// I/O API/IN/STRUCTURE/bds_inPha_measmt_ts
///Data structure for one current measurement value of the API function |bds_inPha_get.|.
{attribute 'external_name' := 'cmp_rts_bds_inPha_measmt_ts'}
TYPE bds_inPha_measmt_ts :
STRUCT
	///Measured current in micro Ampere
	phaShift_dDeg_s32 : DINT;
	///Shunt state of the input current measurement signal
	tiPhaDif_ns_u32: UDINT;
	///Measured current in micro Ampere
	tiPerdPrimSig_ns_u32 : UDINT;
	///Shunt state of the input current measurement signal
	tiPerdSecSig_ns_u32: UDINT;
	///Measured current in micro Ampere
	cntPlsPrimSig_u32 : UDINT;
	///Shunt state of the input current measurement signal
	cntPlsSecSig_u32: UDINT;
	///Shunt state of the input current measurement signal
	statusDiag_b: bds_inPha_statusDiag_tb;
	///Status of the measurement
	status_e: bds_inCmn_status_te;
END_STRUCT
END_TYPE

// I/O API/IN/STRUCTURE/bds_inPha_statusDiag_tb
{attribute 'external_name' := 'cmp_rts_bds_inPha_statusDiag_tb'}
{attribute 'size' := '32'}
TYPE bds_inPha_statusDiag_tb :
STRUCT
	stErrPrimSigMaxPerdOvf_b1: BIT; // Fault error status for maximum period overflow on primary signal;
	stErrSecSigMaxPerdOvf_b1: BIT; // Fault error status for maximum period overflow on secondary signal;
	stErrSigFrqMismatch_b1: BIT; // Fault error status for frequency mismatch of primary and secondary signal.
	resd1_b : ARRAY[0..2] OF BYTE;      (* Reserved *)
END_STRUCT
END_TYPE

// I/O API/IN/STRUCTURE/bds_inPha_tiBufdMeasmt_ts
///Data structure for twenty pwm measurement values of the API function |bds_inPwm_getTiBufd|, used to get the buffered values.
{attribute 'external_name' := 'cmp_rts_bds_inPha_tiBufdMeasmt_ts'}
TYPE bds_inPha_tiBufdMeasmt_ts :
STRUCT
	///Up to 20 samples of PWM period in ns, 0th index is latest
	tiPhaDif_ns_au32: ARRAY[0..19] OF UDINT;
	///Up to 20 samples of ON pulse width in ns
	tiPerdPrimSig_ns_au32: ARRAY[0..19] OF UDINT;
	///Up to 20 samples of ON pulse width in ns
	tiPerdSecSig_ns_au32: ARRAY[0..19] OF UDINT;
	///Number of new samples (pulses) received since the last call of API. It is limited to 20 samples.
	cntPlsPrimSig_u32: UDINT;
	///Number of new samples (pulses) received since the last call of API. It is limited to 20 samples.
	cntPlsSecSig_u32: UDINT;
	///Number of new samples (pulses) received since the last call of API. It is limited to 20 samples.
	cntNewSample_u32: UDINT;
	///Number of new samples (pulses) received since the last call of API. It is limited to 20 samples.
	statusDiag_b: bds_inPha_statusDiag_tb;
END_STRUCT
END_TYPE

// I/O API/IN/STRUCTURE/bds_inPha_tiBufd_ts
///Data structure for pwm measurement value of the API function |bds_inPha_tiBufd_ts|.
{attribute 'external_name' := 'cmp_rts_bds_inPha_tiBufd_ts'}
TYPE bds_inPha_tiBufd_ts :
STRUCT
	///Status of the measurement
	status_e: bds_inCmn_status_te;
END_STRUCT
END_TYPE

// System API/DSM/DSM Refactored( 3-byte DTC)/STRUCTURE/bds_dsmCmn_stWord_tb
///Structure for the Bit field for the 16-bit status word of DFC.
{attribute 'external_name' := 'cmp_rts_bds_dsmCmn_stWord_tb'}
TYPE bds_dsmCmn_stWord_tb :
STRUCT
	///Fault level (0x0 - OK level, 0xF - Defect)
	stFltLvl_b4: BIT;
	///Status of Last Debounced Fault (LDF)
	stLDF_b1: BIT;
	///Tested Since Clear Status (1 - Yes, 0 - No)
	stTSC_b1: BIT;
	///Memory Status (DFC is saved in fault memory or not)
	stMS_b1: BIT;
	///Debounce Active Status (1 - Yes, 0 - No)
	stDA_b1: BIT;
	///Debounced Fault Level (With five levels 0x0, 0x4, 0x8, 0xC and 0xF (e.g., 0xC = 75% debounced)
	stDebdFltLvl_b4: BIT;
	///Fault Since Clear Status (1=Yes, 0=No)
	stFSC_b1: BIT;
	///Test Status
	stTestSt_b1: BIT;
	///Not used
	stUnused_b1: BIT;
	///Test finalized
	stNotFinalized_b1: BIT;
END_STRUCT
END_TYPE

// System API/DSM/DSM Refactored( 3-byte DTC)/STRUCTURE/bds_dsmDTC_deleteErr_ts
///Return structure for bds_dsmDTC_deleteErr POU.
{attribute 'external_name' := 'cmp_rts_bds_dsmDTC_deleteErr_ts'}
TYPE bds_dsmDTC_deleteErr_ts :
STRUCT
	///Status or result of POU operation 
	apiSt_e: bds_dsmCmn_st_te;
END_STRUCT
END_TYPE

// System API/DSM/DSM Refactored( 3-byte DTC)/STRUCTURE/bds_dsmDTC_getDFES_ts
///Return structure for bds_dsmDTC_getDFES POU.
{attribute 'external_name' := 'cmp_rts_bds_dsmDTC_getDFES_ts'}
TYPE bds_dsmDTC_getDFES_ts :
STRUCT
	///Number of errors returned
	nrErr_u8: USINT;
	///DTCs as in DFES array
	dtcListDFES_au32: ARRAY[1..32] OF UDINT;
	///Status or result of POU operation (Valid POU call / Invalid parameter (invalid mask)/ out of Range (DTC value out of range)) 
	apiSt_e: bds_dsmCmn_st_te;
END_STRUCT
END_TYPE

// System API/DSM/DSM Refactored( 3-byte DTC)/STRUCTURE/bds_dsmDTC_getDTCVal_ts
///Return structure for bds_dsmDTC_getDTCVal POU.
{attribute 'external_name' := 'cmp_rts_bds_dsmDTC_getDTCVal_ts'}
TYPE bds_dsmDTC_getDTCVal_ts :
STRUCT
	///DTC value
	dtc_u32: UDINT;
	///Status or result of API operation (API call successful / invalid config (wrong DFC passed) 
	apiSt_e: bds_dsmCmn_st_te;
END_STRUCT
END_TYPE

// System API/DSM/DSM Refactored( 3-byte DTC)/STRUCTURE/bds_dsmDTC_getErrList_ts
///Return structure for bds_dsmDTC_getErrList POU.
{attribute 'external_name' := 'cmp_rts_bds_dsmDTC_getErrList_ts'}
TYPE bds_dsmDTC_getErrList_ts :
STRUCT
	///Number of errors returned
	nrErr_u8: USINT;
	///DTC list containing 32 entries
	dtcList_au32: ARRAY[1..32] OF UDINT;
	///Status or result of POU operation (Valid POU call / Invalid parameter (invalid mask) 
	apiSt_e: bds_dsmCmn_st_te;
END_STRUCT
END_TYPE

// System API/DSM/DSM Refactored( 3-byte DTC)/STRUCTURE/bds_dsmDTC_getStatus_ts
///Return structure for bds_dsmDTC_getStatus POU.
{attribute 'external_name' := 'cmp_rts_bds_dsmDTC_getStatus_ts'}
TYPE bds_dsmDTC_getStatus_ts :
STRUCT
	///Error State (Active / Previously Active / Deactive)
	errState_e: UDINT;
	///DTC Detailed Status Parameters as 16 bit Status Word in DFC
	stWordDTC_b: bds_dsmCmn_stWord_tb;
	///Status or result of POU operation 
	apiSt_e: bds_dsmCmn_st_te;
END_STRUCT
END_TYPE

// System API/DSM/DSM Refactored( 3-byte DTC)/STRUCTURE/bds_dsmDTC_updateErr_ts
///Return structure for bds_dsmDTC_updateErr POU.
{attribute 'external_name' := 'cmp_rts_bds_dsmDTC_updateErr_ts'}
TYPE bds_dsmDTC_updateErr_ts :
STRUCT
	///Status or result of POU operation
	apiSt_e: bds_dsmCmn_st_te;
END_STRUCT
END_TYPE

// Communication API/ISOBUS/J1939-76/STRUCTURE/bds_isobus_cnsrDataboxInfo_ts
///Structure of the consumer data box information
{attribute 'external_name' := 'cmp_rts_bds_isobus_cnsrDataboxInfo_ts'}
TYPE bds_isobus_cnsrDataboxInfo_ts :
STRUCT
	///pointer to the consumer SDG databox buffer
	mem_pas: POINTER TO bds_isobus_cnsrSdgMsg_ts;
	///number of SDG messages to be received
	numOfMsg_u16: UINT;
END_STRUCT
END_TYPE

// Communication API/ISOBUS/J1939-76/STRUCTURE/bds_isobus_cnsrSdgMsg_ts
///Structure for handling Consumer databox
{attribute 'external_name' := 'cmp_rts_bds_isobus_cnsrSdgMsg_ts'}
TYPE bds_isobus_cnsrSdgMsg_ts :
STRUCT
	///pointer to data array with length=lenMax_u8
	data_pau8: POINTER TO USINT;
	///function is called if SDG is received and processed
	func_pf: POINTER TO UINT;
	///CAN Id of the SDM to be received
	canID_u: bds_isobus_sfty_canID_tu;
	///length of received SDM message
	lenAct_u8: USINT;
	///max length of the SDG receive buffer defined
	lenMax_u8: USINT;
	///expected maximum time between consecutive SDMs received
	sct_u32: UDINT;
	///expected maximum time between SHM and SDM of an SDG received
	srvt_u32: UDINT;
	///expected Source address of the sender (i.e., Producer)
	srcAddr_u8: USINT;
	///status of consumer SDG databox
	status_u16: UINT;
	///flag to identify first message received after start-up
	firstSdg_l: BOOL;
	///SCT timer
	sctTmr_s: bds_isobus_sftyTmr_ts;
	///SRVT timer
	srvtTmr_s: bds_isobus_sftyTmr_ts;
	///SDM CRC
	sdmCrc_u: bds_isobus_sdmCrcVal_tu;
	///sequence number handling structure
	seqNum_s: bds_isobus_cnsrSdgSeqNum_ts;
	///SDG state handling enumeration
	sdgState_e: bds_isobus_sdgState_te;
	///Status of Consumer to be updated to ASW
	cnsrStatus_e: bds_isobus_sdgCnsrStatus_te;
END_STRUCT
END_TYPE

// Communication API/ISOBUS/J1939-76/STRUCTURE/bds_isobus_cnsrSdgSeqNum_ts
///Structure type definition for handling CRC32 value of SDM
{attribute 'external_name' := 'cmp_rts_bds_isobus_cnsrSdgSeqNum_ts'}
TYPE bds_isobus_cnsrSdgSeqNum_ts :
STRUCT
	///Sequence number of currently received SDG
	curSdgSeqNum_u8: UINT;
	///Sequence number of previously received SDG, initialize with 0xFF to monitor 0th sequence after start-up
	prevSdgSeqNum_u8: UINT;
END_STRUCT
END_TYPE

// Communication API/ISOBUS/J1939-76/STRUCTURE/bds_isobus_prodDataboxInfo_ts
///Structure of the producer data box information
{attribute 'external_name' := 'cmp_rts_bds_isobus_prodDataboxInfo_ts'}
TYPE bds_isobus_prodDataboxInfo_ts :
STRUCT
	///pointer to the consumer SDG databox buffer
	mem_pas: POINTER TO bds_isobus_prodSdgMsg_ts;
	///number of SDG messages to be transmitted
	numOfMsg_u16: UINT;
END_STRUCT
END_TYPE

// Communication API/ISOBUS/J1939-76/STRUCTURE/bds_isobus_prodSdgMsg_ts
///Structure for handling Producer databox
{attribute 'external_name' := 'cmp_rts_bds_isobus_prodSdgMsg_ts'}
TYPE bds_isobus_prodSdgMsg_ts :
STRUCT
	///pointer to data array updated in Producer callback with length=lenMax_u8
	data_pau8: POINTER TO USINT;
	///function is called before SDG is to be sent (Producer Callback)
	func_pf: POINTER TO UINT;
	///CAN Id of the SDM to be sent
	canID_u: bds_isobus_sfty_canID_tu;
	///max length (buffer size) of SDM to be sent
	lenMax_u8: USINT;
	///actual length of SDM message to be sent
	lenAct_u8: USINT;
	///cycle time for fixed transmission of the SDG
	cycle_u16: UINT;
	///counter for monitoring cyclic transmission of SDG
	counter_u16: UINT;
	///expected Source address of the sender (i.e., Producer)
	srcAddr_u8: USINT;
	///status of Producer SDG databox
	status_u16: UINT;
	///Databox number of the SDG being handled
	SdgDataboxNum_u16: UINT;
	///SDM CRC
	sdmCrc_u: bds_isobus_sdmCrcVal_tu;
	///Sequence number of the SDG being handled
	seqNum_u8: USINT;
	///Timer value of previously transmitted SDG //ToDo: for variable transmission
	prevSdgTmrVal_u32: UDINT;
	///Structure instance containing SHM related data
	shmMsg_s: bds_isobus_shmMsg_ts;
END_STRUCT
END_TYPE

// Communication API/ISOBUS/J1939-76/UNION/bds_isobus_sdmCrcVal_tu
///Union type definition for handling CRC32 value of SDM
{attribute 'external_name' := 'cmp_rts_bds_isobus_sdmCrcVal_tu'}
TYPE bds_isobus_sdmCrcVal_tu :

UNION
	///array containing CRC32 data bytes
	sdmCrcVal_au8: ARRAY[1..4] OF USINT;
	///CRC32 value
	sdmCrcVal_u32: UDINT;
END_UNION

END_TYPE

// Communication API/ISOBUS/J1939-76/STRUCTURE/bds_isobus_sftyTmr_ts
///Structure type definition for Timer handling
{attribute 'external_name' := 'cmp_rts_bds_isobus_sftyTmr_ts_ts'}
TYPE bds_isobus_sftyTmr_ts :
STRUCT
	///timer value for monitoring
	tmrStrd_u32: UDINT;
END_STRUCT
END_TYPE

// Communication API/ISOBUS/J1939-76/STRUCTURE/bds_isobus_sfty_canID_ts
///Structure for handling CAN Id of SHM and SDM.
{attribute 'external_name' := 'cmp_rts_bds_isobus_sfty_canID_ts'}
TYPE bds_isobus_sfty_canID_ts :
STRUCT
	/// node id of the transmitter 
	SourceAddr_b8: BYTE;
	/// if PF<240, this value is destination address else Group extension
	PDUSpecific_b8: BYTE;
	/// this byte determines whether the message can be transmitted with a destination address or as a broadcast
	PDUFormat_b8: BYTE;
	/// these bits identify the data pages of the parameter group
	DataPage_b2: BIT;
	/// these 3 bits define the priority of the following message
	Priority_b3: BIT;
	/// these 3 bits are overhead for the 29 bit CAN Id 
	unusedBits_b3: BIT;
END_STRUCT
END_TYPE

// Communication API/ISOBUS/J1939-76/UNION/bds_isobus_sfty_canID_tu
///Union type definition for handling CAN Id of SHM and SDM
{attribute 'external_name' := 'cmp_rts_bds_isobus_sfty_canID_tu'}
TYPE bds_isobus_sfty_canID_tu :

UNION
	///CAN Id structure of type bds_isobus_sfty_canID_ts
	canID_s: bds_isobus_sfty_canID_ts;
	///CAN Id value
	canID_u32: UDINT;
END_UNION

END_TYPE

// Communication API/ISOBUS/J1939-76/STRUCTURE/bds_isobus_shmMsg_ts
///Structure containing SHM parameters of the bds_isobus_prodSdgMsg_t SDG databox being handled
{attribute 'external_name' := 'cmp_rts_bds_isobus_shmMsg_ts'}
TYPE bds_isobus_shmMsg_ts :
STRUCT
	///array containing CRC32 data bytes
	data_au8: ARRAY[1..8] OF USINT;
	///CAN Id of the SDM to be received
	canID_u: bds_isobus_sfty_canID_tu;
END_STRUCT
END_TYPE

// System API/DSM/DSM Refactored( 3-byte DTC)/ENUM/bds_dsmCmn_st_te
(* common status enumeration return types*)
{attribute 'external_name' := 'cmp_rts_bds_dsmCmn_st_te'}
TYPE bds_dsmCmn_st_te :
(
	(*POU call successful*)
	bds_dsmCmn_ok_E := 0,
	(*Parameter out of Range (e.g., invalid DTC value, which is not within the configured Range)*)
	bds_dsmCmn_outOfRng_E,
	(*not available (e.g. busy, called to early in init, System in a mode it cannot measure etc.)*)
    bds_dsmCmn_notAvl_E,
	(*POU call invalid, e.g., calling a not configured DFC, etc.*)
    bds_dsmCmn_invldCfg_E,
	(*POU call invalid because of invalid Parameter*)
    bds_dsmCmn_invldPrm_E,
	(*POU call invalid because of invalid pointer*)
    bds_dsmCmn_invldPtr_E,
	(*Not available due to an internal error*)
    bds_dsmCmn_errInt_E
	
)USINT;
END_TYPE

// System API/DSM/DSM Refactored( 3-byte DTC)/ENUM/bds_dsmCmn_errState_te
(*Enumeration containing the error state of DFC (Active / Previously Active / Deactive).*)
{attribute 'external_name' := 'cmp_rts_bds_dsmCmn_errState_te'}
TYPE bds_dsmCmn_errState_te :
(
	(*Error is Active*)
	bds_dsmCmn_stErrActv_e := 1,
	(*Error is Previously Active*)
	bds_dsmCmn_stErrPrevActv_e,
	(*Error is in Deactive State*)
	bds_dsmCmn_stErrDeactv_e
	
)USINT;
END_TYPE

// System API/DSM/DSM Refactored( 3-byte DTC)/ENUM/bds_dsmCmn_fltLvl_te
(*Enumeration for fault level of a DFC, as a result of check.*)
{attribute 'external_name' := 'cmp_rts_bds_dsmCmn_fltLvl_te'}
TYPE bds_dsmCmn_fltLvl_te :
(
	(*Fault percent 0%*)
	bds_dsmCmn_fltLvl_0_Perc_e := 0,
	(*Fault percent 100%*)
	bds_dsmCmn_fltLvl_100_Perc_e
	
)USINT;
END_TYPE

// System API/DSM/DSM Refactored( 3-byte DTC)/STRUCTURE/bds_dsmJ1939_LampSt_tb
(*Bit field for Lamp States.*)
{attribute 'external_name' := 'cmp_rts_bds_dsmJ1939_LampSt_tb'}
TYPE bds_dsmJ1939_LampSt_tb :
STRUCT
	(*Lamp/Flash State of Malfunction Indicator Lamp (MIL)*)
	milSt_b2: BIT;
	(*Lamp/Flash State of Red Stop Lamp (RSL)*)
	rslSt_b2: BIT;
	(*Lamp/Flash State of Amber Warning Lamp (AWL)*)
	awlSt_b2: BIT;
	(*Lamp/Flash State of Protected Lamp (PRL)*)
	prlSt_b2: BIT;
END_STRUCT
END_TYPE

// System API/DSM/DSM Refactored( 3-byte DTC)/STRUCTURE/bds_dsmJ1939_getJ1939DTC_ts
(*Return structure for the bds_dsmJ1939_getJ1939DTC POU.*)
{attribute 'external_name' := 'cmp_rts_bds_dsmJ1939_getJ1939DTC_ts'}
TYPE bds_dsmJ1939_getJ1939DTC_ts :
STRUCT
	(*SPN value*)
	spn_u32 : UDINT;
	(*FMI value*)
	fmi_u8 : USINT;
	(*Bitfield containing Lamp States (MIL, RSL, AWL, Protected Lamp)*)
	lampSt_b : bds_dsmJ1939_LampSt_tb;
	(*Occurrence Counter*)
	occCntr_u8 : USINT;
	(* Status or result of POU operation (Valid POU call / DTC passed is out of range)*)
	apiSt_e : bds_dsmCmn_st_te;
END_STRUCT
END_TYPE

// Communication API/CAN/CAN-FD legacy/ENUM/bds_can_fd_St_te
{attribute 'external_name' := 'cmp_rts_bds_can_fd_St_te'}
TYPE bds_can_fd_St_te :
(
	//API call successful
    bds_can_fd_ok_E := 0,
	//Databox not empty
    bds_can_fd_txDataboxNotEmpty_E := 1,
	//Invalid Access to FFI variant API call.
    bds_can_fd_errFfi_E := 5,
	//Invalid CAN-FD databox number
    bds_can_fd_invldDataBoxNbr_E := 9,
	//Invalid CAN-FD channel
    bds_can_fd_invldChnl_E := 14,
	//Invalid CAN-FD identifier
    bds_can_fd_invldId_E := 15,
	//Invalid CAN-FD message format
    bds_can_fd_invldFormat_E := 16,
	//Invalid number of bytes
    bds_can_fd_invldNumBytes_E := 17,
	//Number of messages registered in buffer = 0
    bds_can_fd_numMsgZero_E := 18,
	//CAN-FD transmit buffer overflow
    bds_can_fd_txBufOvfl_E := 20,
	//CAN-FD receive buffer overflow
    bds_can_fd_rxBufOvfl_E := 30,
	//CAN-FD receive buffer is empty
    bds_can_fd_rxBufEmpty_E := 31,
	//CAN-FD receive buffer length is zero
    bds_can_fd_rxBufLenZero_E := 32,
	//Buffer address overlap
    bds_can_fd_ovlpAddr_E := 55,
	//Invalid address
    bds_can_fd_invldAddr_E := 60,
	//Invalid address (parameter buf_pas). Buffer length is zero
    bds_can_fd_rxDataboxBufLenZero_E := 61,
	//Databox not initialized
    bds_can_fd_dataBoxNoInit_E := 62,
	//Databox with this identifier is initialized already, new initialization is not accepted
    bds_can_fd_errDataboxIdExist_E := 63,
	//Number of databoxes registered is greater than previously registered number of databoxes
    bds_can_fd_prevRegdDataboxMoreThanCurrent_E := 64,
	//Invalid number of databoxes
    bds_can_fd_invldCfgDatabox_E := 65,
	//CAN hardware not supported in RC.
    //e.g., 3 CAN channel RC5-6/40 ECU.
    bds_can_fd_hwNotSupported_E := 66,
	//Configuration not allowed
    bds_can_fd_cfgNotAllowed_E := 99,
	//CAN-FD not supported in CAN_3
    bds_can_fd_paramChnl3Err_E := 100
)USINT;
END_TYPE

// Communication API/CAN/CAN-FD legacy/STRUCTURE/bds_can_fd_Message_ts
{attribute 'external_name' := 'cmp_rts_bds_can_fd_Message_ts'}
TYPE bds_can_fd_Message_ts :
STRUCT
	//Identifier of the message.
	//Value range:
	// 16#000 .. 0x7FF (11-bit standard format)
	// 16#00000000 .. 0x1FFFFFFF (29-bit extented format)
	id_u32 : UDINT;
	//Format of the CAN-FD message.Value range:
    //BDS_CAN_STD_DU8 (11-bit standard format)
	//BDS_CAN_EXD_DU8 (29-bit extented format)
	format_u8 : USINT;
	//Number of data bytes which will be transmitted or which type received.
	numBytes_u8 : USINT;
	//Data which will be transmitted or which were received.Size of the define, bds_can_fd_maxDataBytes_DU8 is equal to 64.
	data_au8 : ARRAY[0..63] OF USINT;
END_STRUCT
END_TYPE

// Communication API/ISOBUS/J1939-76/ENUM/bds_isobus_sdgCnsrStatus_te
(*Enumeration for Consumer SDG reception status.*)
{attribute 'external_name' := 'cmp_rts_bds_isobus_sdgCnsrStatus_te'} 
TYPE  bds_isobus_sdgCnsrStatus_te :
(  
	(*valid SDG received*)
	bds_isobus_sdgCnsrOk_E := 0,
	(*SRVT timeout*)
	bds_isobus_sdgCnsrSrvtTmngErr_E,
	(*SCT timeout*)
	bds_isobus_sdgCnsrSctTmngErr_E,
	(*SDG received with invalid CRC*)
    bds_isobus_sdgCnsrCrcError_E,
	(*SDG received with invalid sequence number*)
    bds_isobus_sdgCnsrSeqError_E,
	(*SDG received with invalid data length*)
    bds_isobus_sdgCnsrLenError_E
)USINT;
END_TYPE

// Communication API/ISOBUS/J1939-76/ENUM/bds_isobus_sdgState_te
(*Enumeration for Consumer SDG reception status.*)
{attribute 'external_name' := 'cmp_rts_bds_isobus_sdgState_te'} 
TYPE bds_isobus_sdgState_te :
(
	(*SDG initialized*)
	bds_isobus_sfty_sdgIniDone_E := 0,
	(*SHM received and processed*)
	bds_isobus_sfty_shmProcessed_E,
	(*both SHM and SDM received and processed*)
	bds_isobus_sfty_sdgProcessed_E,
	(*SRVT timeout*)
	bds_isobus_sfty_srvtExpired_E,
	(*SCT timeout*)
	bds_isobus_sfty_sctExpired_E,
	(*SDG successfully validated*)
	bds_isobus_sfty_sdgValidated_E,
	(*Consumer SDG callback triggered*)
	bds_isobus_sfty_cnsrSdgCbkTriggered_E
)USINT;
END_TYPE

// Communication API/ISOBUS/J1939-76/ENUM/bds_isobus_sfty_apiRetVal_te
(*Enumeration for J1939-76 API return values.*)
{attribute 'external_name' := 'cmp_rts_bds_isobus_sfty_apiRetVal_te'}
TYPE bds_isobus_sfty_apiRetVal_te :
(
	(*No API execution error*)
	 bds_isobus_sfty_noErr_E := 0,
	(*invalid address*)
	 bds_isobus_sfty_invldAdr_E,
	(*address overlaps with other buffers*)
 	 bds_isobus_sfty_ovlAdr_E,
	(*invalid CA instance number*)
	 bds_isobus_sfty_invldInstNum_E,
	(*message box is not yet initialized*)
	 bds_isobus_sfty_boxStNoIni_E,
	(*configuration is not allowed*)
	 bds_isobus_sfty_boxStIni_E,
	(*invalid databox number*)
	 bds_isobus_sfty_cfgNotAllwd_E,
	(*invalid PGN value*)
	 bds_isobus_sfty_invldDataboxNum_E,
	(* invalid priority of SDG*) 
	 bds_isobus_sfty_invldPgn_E,
	(*invalid cycle time for SDG*)
	 bds_isobus_sfty_invldPrio_E,
	(*invalid offset time for SDG*)
	 bds_isobus_sfty_invldCyc_E,
	(*invalid data length of SDM*)
	 bds_isobus_sfty_invldOffs_E,
	(*invalid data address*)
	 bds_isobus_sfty_invldDataLen_E,
	(*Another data box with this id was initialized already*) 
	 bds_isobus_sfty_invldDataPtr_E,
	(*sdg databox initialized*) 
	 bds_isobus_sfty_pgnPrioExists_E,
	(*invalid source address*)
	 bds_isobus_sfty_invldSrcAdr_E,
	(*invalid SCT*)
	 bds_isobus_sfty_invldSct_E,
	(*invalid SRVT*) 
	 bds_isobus_sfty_invldSrvt_E,
	(*Internal PGN used*) 
	 bds_isobus_sfty_intPgnUsed_E,
	(*API used without enabling J1939-76 feature in eC*)
	 bds_isobus_sfty_featNotEnad_E,
	(*Invalid pointer*)
	 bds_isobus_sfty_invldCbkAdr_E
)USINT;
END_TYPE

// Diagnostics API/UDS/ENUM/bds_udsCmn_statusApi_te
{attribute 'external_name' := 'cmp_rts_bds_udsCmn_statusApi_te'}
TYPE bds_udsCmn_statusApi_te :
(
	(*Success: API executed without error*)
	bds_udsCmn_ok_E := 0,
	(*Invalid: calling an unconfigured signal/DID *)
	bds_udsCmn_invldCfg_E,
	(*Invalid: invalid parameter*)
	bds_udsCmn_invldPrm_E,
	(*Out of range: the array size should be less than or equal to 17 bytes*)
	bds_udsCmn_outOfRng_E,
	(*not available: (e.g. busy, called to early in init, system is in a mode that it cannot measure etc)*)
	bds_udsCmn_notAvl_E
)USINT;
END_TYPE

// Communication API/CAN/CAN-FD legacy/STRUCTURE/bds_can_fd_RxDatabox_ts
///Structure of a CAN-FD receive (Rx) databox.
{attribute 'external_name' := 'cmp_rts_bds_can_fd_RxDatabox_ts'}
TYPE bds_can_fd_RxDatabox_ts :
STRUCT
	//CAN ID
    //Value range:
    //16#000 .. 0x7FF (11-bit standard format)
    // 16#00000000 .. 16#1FFFFFFF (29-bit extented format)
	id_u32 : UDINT;
	//CAN ID format
    //Value range:
    //BDS_CAN_STD_DU8 (11-bit standard format)
    //BDS_CAN_EXD_DU8 (29-bit extented format)
	format_u8 : USINT;
	//Number of data bytes which will be received.
    numBytes_u8 : USINT;
	//Pointer to callback function for CAN-FD Receive Databox
    callback_pf : UINT;
	//Structure instance to CAN-FD databox buffer information
    Buf_s : bds_can_fd_DataboxBufInfo_ts;
END_STRUCT
END_TYPE

// Communication API/CAN/CAN-FD legacy/STRUCTURE/bds_can_fd_DataboxData_ts
///Structure of data of a CAN-FD databox.
{attribute 'external_name' := 'cmp_rts_bds_can_fd_DataboxData_ts'}
TYPE bds_can_fd_DataboxData_ts :
STRUCT
	//Received data.Size of the define, bds_can_fd_maxDataBytes_DU8 is equal to 64.
	data_au8 : ARRAY[0..63] OF USINT;
	//Number of data bytes received
	numBytes_u8 : USINT;
END_STRUCT
END_TYPE

// Communication API/CAN/CAN-FD legacy/STRUCTURE/bds_can_fd_DataboxBufInfo_ts
///Structure for a CAN-FD databox buffer. Only data of the CAN-FD message is buffered.
{attribute 'external_name' := 'cmp_rts_bds_can_fd_DataboxBufInfo_ts'}
TYPE bds_can_fd_DataboxBufInfo_ts :
STRUCT
	//Pointer to structure for CAN-FD Databox Data structure.
	start_pas : POINTER TO bds_can_fd_DataboxData_ts;
	//CAN-FD Databox Buffer Management Structure 
	Manage_s : bds_can_fd_BufManage_ts;
END_STRUCT
END_TYPE

// Communication API/CAN/CAN-FD legacy/STRUCTURE/bds_can_fd_BufManage_ts
///Structure for a CAN-FD Message Buffer Management.
{attribute 'external_name' := 'cmp_rts_bds_can_fd_BufManage_ts'}
TYPE bds_can_fd_BufManage_ts :
STRUCT
	//Length of the buffer
	length_u16 : UINT;
	//Index for write (CAN-FD send / receive) in the buffer.This is for buffer (FIFO - in sequence value).
	//This is more specific to BSW, has lesser significance to application.
	idx_in_u16 : UINT;
	//Index for read (CAN-FD send / receive) out of the buffer.This is for buffer ((FIFO - out sequence value).
	//This is more specific to BSW, has lesser significance to application.
    idx_out_u16 : UINT;
	//FALSE: Buffer is not empty. If then idx_out - idx_in: buffer is full (no put in).
    //TRUE: Buffer is empty (nothing is to send or nothing was received)
	BufEmpty_l : BOOL;
	//This flag shows if a buffer overflow is occurred.
	//FALSE: No buffer overflow is occurred since last user inquiry of status
    //TRUE: Buffer overflow is occurred.
    BufOvfl_l : BOOL;
END_STRUCT
END_TYPE

// Communication API/CAN/CAN-FD legacy/STRUCTURE/bds_can_fd_TxDatabox_ts
///Structure of a CAN-FD transmit (Tx) databox.
{attribute 'external_name' := 'cmp_rts_bds_can_fd_TxDatabox_ts'}
TYPE bds_can_fd_TxDatabox_ts :
STRUCT
	//CAN ID
    //Value range:
    //16#000 .. 0x7FF (11-bit standard format)
    // 16#00000000 .. 16#1FFFFFFF (29-bit extented format)
	id_u32 : UDINT;
	//CAN ID format
    //Value range:
    //BDS_CAN_STD_DU8 (11-bit standard format)
    //BDS_CAN_EXD_DU8 (29-bit extented format)
	format_u8 : USINT;
	//Number of data bytes which will be received.
    numBytes_u8 : USINT;
	//Data which will be transmitted or which were received.Size of the define, bds_can_fd_maxDataBytes_DU8 is equal to 64.
	data_au8 : ARRAY[0..63] OF USINT;
	//TRUE = databox is empty
    //FALSE = databox contains data which were not sent
    empty_l : BOOL;
	//TRUE = databox is initialized
    //FALSE = databox is not yet initialized
    init_l : BOOL;
END_STRUCT
END_TYPE

// Communication API/ISOBUS/STRUCTURE/bds_isobus_caAddrInfoTbl_ts
///Structure definition of an ISOBUS address info table.
{attribute 'external_name' := 'cmp_rts_bds_isobus_caAddrInfoTbl_ts'}
TYPE bds_isobus_caAddrInfoTbl_ts :
STRUCT
	//ISOBUS CA Name, which is 8 bytes in size according to the ISOBUS/J1939 specification.
	caName_au8 : ARRAY[0..7] OF USINT;
	//ISOBUS CA address which is 1 byte in size.
	caAddr_u8 : USINT;
END_STRUCT
END_TYPE

// Diagnostics API/UDS/STRUCTURE/bds_uds_getActiveService_ts
///Return structure for the API function bds_uds_getActiveService.
{attribute 'external_name' := 'cmp_rts_bds_uds_getActiveService_ts'}
TYPE bds_uds_getActiveService_ts :
STRUCT
	//Status of the UDS API function call.
	stsApi_e : bds_udsCmn_statusApi_te;
	//The value of the UDS service identifier.
    dataSid_u8 : USINT;
END_STRUCT
END_TYPE

// Communication API/ISOBUS/ENUM/bds_isobus_caAddrCbEventType_te
{attribute 'external_name' := 'cmp_rts_bds_isobus_caAddrCbEventType_te'}
TYPE bds_isobus_caAddrCbEventType_te :
(
	//Address claim message received, address table entry is not updated
	bds_isobus_addrClaimMsgRcv_E := 0,
	//Address claim message received and address table entry is updated with new address
    bds_isobus_caTbleAddressUpdate_E,
	//Address claim message received and new entry created in address table
	bds_isobus_caTbleNewEntry_E
)USINT;
END_TYPE

// Communication API/ISOBUS/STRUCTURE/bds_isobus_caAddrInfoTblRef_ts
//Structure type definition to hold reference to Address table info and size of address table info
{attribute 'external_name' := 'cmp_rts_bds_isobus_caAddrInfoTblRef_ts'}
TYPE bds_isobus_caAddrInfoTblRef_ts :
STRUCT
	//pointer to Address Info table
	mem_pas : POINTER TO bds_isobus_caAddrInfoTbl_ts;
	//Total number (Size) of Entries in address info table
	numOfEntry_u8 : USINT;
	//Last valid entry/Number of valid entries in address info table
	lastEntry_u8 : USINT;
END_STRUCT
END_TYPE

// Communication API/Ethernet/STRUCTURE/bds_ethIPv4_getLocalIpAdr_ts
{attribute 'external_name' := 'cmp_rts_bds_ethIPv4_getLocalIpAdr_ts'}
TYPE bds_ethIPv4_getLocalIpAdr_ts :
STRUCT
	//The return structure containing the status information
	statusApi_e : bds_ethIPv4_statusApi_te; 
END_STRUCT
END_TYPE

// Communication API/Ethernet/ENUMS/bds_ethIPv4_statusApi_te
{attribute 'external_name' := 'cmp_rts_bds_ethIPv4_statusApi_te'}
TYPE bds_ethIPv4_statusApi_te :
(
	//API call is successful
	bds_ethIPv4_Adr_Mask_ok_E := 0,
	//API call is invalid because of invalid IPv4 address
    bds_ethIPv4_Adr_Nok_E := 1,
	//API call is invalid because of invalid subnet mask, subnet mask should be 16
    bds_ethIPv4_Mask_Nok_E := 2,
	//Not Available (e.g. busy, called too early in init, not called from OsIniProc etc.)
    bds_ethIPv4_Api_NotAvailable_E := 3, 
	//Invalid parameter passed
    bds_ethIPv4_NullPtr_E := 4, 
    bds_ethIPv4_notAssigned_E :=5 
)USINT;
END_TYPE

// Communication API/Ethernet/STRUCTURE/bds_ethIPv4_setLocalIpAdr_ts
{attribute 'external_name' := 'cmp_rts_bds_ethIPv4_setLocalIpAdr_ts'}
TYPE bds_ethIPv4_setLocalIpAdr_ts :
STRUCT
	//The return structure containing the status information
	statusApi_e : bds_ethIPv4_statusApi_te; 
END_STRUCT
END_TYPE

// Communication API/Ethernet/STRUCTURE/bds_ethIPv4_LocalIpAdr_ts
//Data Structure for IPv4 Address and Subnet Mask for Ethernet functions - bds_ethIPv4_setLocalIpAdr and bds_ethIPv4_getLocalIpAdr
{attribute 'external_name' := 'cmp_rts_bds_ethIPv4_LocalIpAdr_ts'}
TYPE bds_ethIPv4_LocalIpAdr_ts :
STRUCT
	//4 bytes of IPv4 Address
	Ipv4Adr_u32 : UDINT;
	//1 byte of Subnet Mask for IPv4
	Ipv4SubnetMask_u8 : USINT;
END_STRUCT
END_TYPE

// Communication API/Ethernet/ENUMS/bds_ethIPv4_linkState_te
//This enum defines the return values for API bds_ethIPv4_setDoipAdr.
{attribute 'external_name' := 'cmp_rts_bds_ethIPv4_linkState_te'}
TYPE bds_ethIPv4_linkState_te :
(
	bds_ethIPv4_linkDown_E := 0,
	bds_ethIPv4_linkUp_E := 1,
	bds_ethIPv4_linkUndef_E
)USINT;
END_TYPE

// Communication API/Ethernet/ENUMS/bds_ethIPv4_retDoipAdr_te
//This enum defines the return values for API bds_ethIPv4_setDoipAdr.
{attribute 'external_name' := 'cmp_rts_bds_ethIPv4_retDoipAdr_te'}
TYPE bds_ethIPv4_retDoipAdr_te :
(
	//Address set successfully 
	bds_ethIPv4_retAdrOk_E := 0,
	//RC4x Logical Address out of range
	bds_ethIPv4_retLogAdrNok_E :=1,
	//Tester Address out of range
	bds_ethIPv4_retTesterAdrNok_E :=2,
	//ECU and Tester Addresses are equal
	bds_ethIPv4_retAdrSame_E :=3,
	//API called outside of OsIniProc
	bds_ethIPv4_retApiNA_E :=4
)USINT;
END_TYPE

// Communication API/Ethernet/ENUMS/bds_ethIPv4_retLinkState_te
{attribute 'external_name' := 'cmp_rts_bds_ethIPv4_retLinkState_te'}
TYPE bds_ethIPv4_retLinkState_te :
(
	//Link status retrieved successfully
	bds_ethIPv4_retLinkOk_E := 0,
	//Failed to get link status
	bds_ethIPv4_retLinkNok_E :=1,
	//Invalid parameter - NULL pointer passed as argument
	bds_ethIPv4_retLinkNull_E :=2
)USINT;
END_TYPE

// Communication API/Ethernet/STRUCTURE/bds_ethIPv4_linkStateInfo_ts
{attribute 'external_name' := 'cmp_rts_bds_ethIPv4_linkStateInfo_ts'}
TYPE bds_ethIPv4_linkStateInfo_ts :
STRUCT
	//Current state of the Ethernet link (up/down/undefined)
	currentState_e : bds_ethIPv4_linkState_te;
END_STRUCT
END_TYPE

// Diagnostics API/UDS/ENUM/bds_uds_setNodeIdTesterId_te
{attribute 'external_name' := 'cmp_rts_bds_uds_setNodeIdTesterId_te'}
TYPE bds_uds_setNodeIdTesterId_te :
(
	//Node Id and Tester Id is set.
	bds_uds_nodeIdTesterIdOk_E := 0,
	//0xFF is broadcast node ID which cannot be used
	bds_uds_nodeIdNotOk_E := 1,
	//0xFF is broadcast tester ID which cannot be used
	bds_uds_testerIdNotOk_E := 2,
	//Node ID and tester ID value cannot be same.
	bds_uds_sameNodeIdTesterIdNotOk_E := 3,
	//This API shall be called from initialization task and cannot be called from elsewhere
 	bds_uds_setIdApiNotAvailable_E := 4
);
END_TYPE

// System API/SYS/ENUM/bds_sys_regOverwriteOpHrs_te
{attribute 'external_name' := 'cmp_rts_bds_sys_regOverwriteOpHrs_te'}
TYPE bds_sys_regOverwriteOpHrs_te :
(
//Callback function registered successfully 
 bds_sys_regOpHrsOk_E := 0,
//A null pointer error occurred for the callback.
 bds_sys_regOpHrsNullPtr_E := 1,
//The API is only available from OsIniProc and cannot be called from elsewhere. 
 bds_sys_regOpHrsApiNotAvailable_E := 2
)USINT;
END_TYPE

// Communication API/CAN/GVL/GVL_can
VAR_GLOBAL
	CANIF_CS_UNINIT: UINT := 0;
	CANIF_CS_STOPPED: UINT := 1;
	CANIF_CS_STARTED: UINT := 2;
	CANIF_CS_SLEEP: UINT := 3;
	///standard 11 bit CAN id
	BDS_CAN_STD_DU8: USINT := 0;
	///extended 29 bit CAN id
	BDS_CAN_EXD_DU8: USINT := 1;
	///flexible data rate with standard 11 bit CAN id
	BDS_CAN_STD_FD_DU8: USINT := 2;
	///flexible data rate with extended 29 bit CAN id
	BDS_CAN_EXD_FD_DU8: USINT := 3;
	BDS_CAN_STD_MAX_ID_DU32: UDINT := 16#7FF;
	BDS_CAN_EXD_MAX_ID_DU32: UDINT := 16#1FFFFFFF;
	BDS_CAN_NONE_ID_DU32: UDINT := 16#FFFFFFFF;
	BDS_CAN_DATALEN_08_DU8: USINT := 8;
	BDS_CAN_DATALEN_12_DU8: USINT := 12;
	BDS_CAN_DATALEN_16_DU8: USINT := 16;
	BDS_CAN_DATALEN_20_DU8: USINT := 20;
	BDS_CAN_DATALEN_24_DU8: USINT := 24;
	BDS_CAN_DATALEN_32_DU8: USINT := 32;
	BDS_CAN_DATALEN_48_DU8: USINT := 48;
	BDS_CAN_DATALEN_64_DU8: USINT := 64;
	BDS_CAN_MAX_STD_DATA_DU8: USINT := BDS_CAN_DATALEN_08_DU8;
	BDS_CAN_MAX_FD_DATA_DU8: USINT := BDS_CAN_DATALEN_64_DU8;
	BDS_CAN_MAX_FD_LEN_D: USINT := 10;
	BDS_CAN_MAX_MSG_SIZE_DU8: USINT := BDS_CAN_MAX_STD_DATA_DU8;
	BDS_BAUD_2000K_DU32: UDINT := 2000000;
	BDS_BAUD_1000K_DU32: UDINT := 1000000;
	BDS_BAUD_500K_DU32: UDINT := 500000;
	BDS_BAUD_250K_DU32: UDINT := 250000;
	BDS_BAUD_125K_DU32: UDINT := 125000;
	BDS_BAUD_100K_DU32: UDINT := 100000;
	BDS_CAN_ERR_NO_ERRORS_DU16: UINT := 0;
	BDS_CAN_ERR_UNKNOWN_BAUDRATE_DU16: UINT := 1;
	///invalid sample point
	BDS_CAN_ERR_SAMPLEPOINT_DU16: UINT := 2;
	///invalid buffer type
	BDS_CAN_ERR_INV_BUF_TYPE_DU16: UINT := 2;
	///invalid CAN FD baudrate
	BDS_CAN_ERR_FD_BAUDRATE_DU16: UINT := 3;
	///Data box number is invalid.
	BDS_CAN_ERR_DATABOXNUM_DU16: UINT := 9;
	///invalid channel (node)
	BDS_CAN_ERR_CHNL_DU16: UINT := 14;
	///invalid id
	BDS_CAN_ERR_ID_DU16: UINT := 15;
	///invalid format
	BDS_CAN_ERR_FORMAT_DU16: UINT := 16;
	///invalid number of data bytes
	BDS_CAN_ERR_NUM_DATA_DU16: UINT := 17;
	///invalid number of messages
	BDS_CAN_ERR_NUM_MSG_DU16: UINT := 18;
	///invalid mask
	BDS_CAN_ERR_MASK_DU16: UINT := 19;
	///Transmit buffer overflow
	BDS_CAN_ERR_TXBUF_OVFL_DU16: UINT := 20;
	///Receive buffer overflow.
	BDS_CAN_ERR_RXBUF_OVFL_DU16: UINT := 30;
	///Receive buffer is empty.
	BDS_CAN_ERR_RXBUF_EMPTY_DU16: UINT := 31;
	///Receive buffer length is zero.
	BDS_CAN_ERR_RXBUF_LEN0_DU16: UINT := 32;
	///A buffer which has to be registered by application(with the help of can-API functions) overlaps with a present buffer registered by application.
	BDS_CAN_ERR_OVERLAP_ADDR_DU16: UINT := 55;
	///Invalid address.
	BDS_CAN_ERR_INVALID_ADDR_DU16: UINT := 60;
	///Buffer length of a databox is zero.
	BDS_CAN_ERR_DATABOX_BUFLEN0_DU16: UINT := 61;
	/// Data box is not initialised.
	BDS_CAN_ERR_DATABOX_NOINIT_DU16: UINT := 62;
	///A data box with this id is initialised already.
	BDS_CAN_ERR_DATABOX_ID_EXIST_DU16: UINT := 63;
	///Number of databoxes registered already is greater
	///than the new number.
	BDS_CAN_ERR_DATABOXES_NUM_OLD_NEW_DU16: UINT := 64;
	///invalid number of databoxes
	BDS_CAN_ERR_DATABOXES_NUM_DU16: UINT := 65;
	///Configuration is not allowed.
	BDS_CAN_ERR_CFG_NOTALLOWED_DU16: UINT := 99;
	///I-PDU group vector address invalid
	BDS_CANSIG_ERR_NULLIPDUVECTOR_DU16: UINT := 110;
	///Initialization parameter invalid
	BDS_CANSIG_ERR_BITFLAG_DU16: UINT := 111;
	///Invalid Tx signal Id
	BDS_CANSIG_ERR_NUM_TX_SIG_DU16: UINT := 112;
	///Invalid Rx signal Id
	BDS_CANSIG_ERR_NUM_RX_SIG_DU16: UINT := 113;
	///Invalid Tx signal Data pointer
	BDS_CANSIG_ERR_TX_DATAPTR_DU16: UINT := 114;
	///Invalid Rx signal Data pointer
	BDS_CANSIG_ERR_RX_DATAPTR_DU16: UINT := 115;
	///Invalid Rx signal length pointer
	BDS_CANSIG_ERR_RX_LENPTR_DU16: UINT := 116;
	///Signal Transmission failure
	BDS_CANSIG_ERR_TX_FAIL_DU16: UINT := 117;
	///Signal Reception failure
	BDS_CANSIG_ERR_RX_FAIL_DU16: UINT := 118;
	///Tx I-PDU not ready
	BDS_CANSIG_ERR_TX_NOSERVICE_DU16: UINT := 119;
	///Rx I-PDU not ready
	BDS_CANSIG_ERR_RX_NOSERVICE_DU16: UINT := 120;
	///Tx databox is empty
	BDS_CAN_TX_DATABOX_EMPTY_DU16: UINT := 0;
	///Tx databox is not empty
	BDS_CAN_TX_DATABOX_NOT_EMPTY_DU16: UINT := 1;
	///Transmitter is empty
	BDS_CAN_TX_CHANNEL_EMPTY_DU16: UINT := 0;
	///Transmitter is not empty
	BDS_CAN_TX_CHANNEL_NOT_EMPTY_DU16: UINT := 1;
	///Invalid CAN channel
	BDS_CAN_TX_CHANNEL_INV_CAN_DU16: UINT := 2;
	/// bit 0: buffer
	BDS_CAN_BUFTYPE_BUF_DU8: USINT := 16#1;
	///bit 1: data boxes
	BDS_CAN_BUFTYPE_DATABOXES_DU8: USINT := 16#2;
	BDS_CAN_STATE_UNINIT_DU16: UINT := CANIF_CS_UNINIT;
	BDS_CAN_STATE_STOPPED_DU16: UINT := CANIF_CS_STOPPED;
	BDS_CAN_STATE_STARTED_DU16: UINT := CANIF_CS_STARTED;
	BDS_CAN_STATE_SLEEP_DU16: UINT := CANIF_CS_SLEEP;
	BDS_CAN_NUM_NODE_D: USINT := 4;
	BDS_CAN_ERR_HW_NOT_SUPPORTED_DU16: UINT := 66;
	BDS_CAN_FFI_ACCESS_ERROR_DU16: UINT := 5;
END_VAR

// System API/DSM/GVL/GVL_dsm
VAR_GLOBAL
	BDS_DSM_ERR_TESTERROR_NOTACTIVE_DU8: USINT := 0;
	BDS_DSM_ERR_TESTERROR_ACTIVE_DU8: USINT := 1;
	///MASK for the DFC
	BDS_DSM_SET_ACTIVE_ERROR_MASK_DU16: UINT := 16#18;
	///MASK for the DFC
	BDS_DSM_SET_TESTED_ONCE_MASK_DU16: UINT := 16#8;
	///MASK for the DFC
	BDS_DSM_SET_TESTED_OK_MASK_DU16: UINT := 16#20;
	///MASK for the DFC
	BDS_DSM_SET_FAILED_SINCE_CLEAR_MASK_DU16: UINT := 16#80;
	///Mask for DFC status
	BDS_DSM_STATUS_ACTIVE_MASK_DU8: USINT := 16#1;
	///Mask for DFC status
	BDS_DSM_STATUS_PREVIOUSLY_ACTIVE_MASK_DU8: USINT := 16#2;
	///Mask for DFC status
	BDS_DSM_STATUS_DEACTIVE_MASK_DU8: USINT := 16#4;
	///Mask for DFC status
	BDS_DSM_STATUS_TESTED_SINCE_CLEAR_MASK_DU8: USINT := 16#8;
	///Mask for DFC status
	BDS_DSM_STATUS_FAULT_SINCE_CLEAR_MASK_DU8: USINT := 16#10;
	BDS_DSM_FAULT_PERCENT_00_DU8: USINT := 0;
	BDS_DSM_FAULT_PERCENT_100_DU8: USINT := 15;
	BDS_DSM_ERR_PERMISSION_DU8: USINT := 0;
	BDS_DSM_ERR_NO_PERMISSION_DU8: USINT := 1;
	BDS_DSM_NO_ERROR_DU16: UINT := 0;
	BDS_DSM_DEBOUNCE_ERROR_DU16: UINT := 2;
	BDS_DSM_DFC_ERROR_DU16: UINT := 1;
	BDS_DSM_NO_DEBOUNCE_ERROR_DU16: UINT := 2;
	BDS_DSM_FAULT_PERCENT_ERROR_DU16: UINT := 3;
	BDS_DSM_INVALID_PTR_DU16: UINT := 4;
	BDS_DSM_MASK_ERROR_DU16: UINT := 5;
	BDS_DSM_MASK_PENDING_DU16: UINT := 6;
	BDS_DSM_INVALID_MAX_ERROR_DU16: UINT := 7;
	BDS_DSM_OVERFLOW_ERROR_DU16: UINT := 8;
	BDS_DSM_NO_DTC_AVAILABLE_DU16: UINT := 11;
	BDS_DSM_WRONG_BUFFERSIZE_DU16: UINT := 10;
	BDS_DSM_DFC_NOEXIST_DU16: UINT := 9;
	BDS_DSM_FFI_ACCESS_ERROR_DU16: UINT := 12;
	///DSM Refactored 3-byte DTC
	bds_dsmCmn_setActvErrMsk_DU16: UINT := 16#18;
	///DFC was tested at least once since start or reset as per DFC status
	bds_dsmCmn_tstdOnceMsk_DU16: UINT := 16#8;
	///DFC was at least once OK tested since start or reset according to status of DFC
	bds_dsmCmn_setTstdOkMsk_DU16: UINT := 16#20;
	///Fault occured at least once since error was detected from memory, with respect to the status of DFC. 
	bds_dsmCmn_setFailedClrMsk_DU16: UINT := 16#80;
	///Buffer size of error List (DTCs/DFCs) for a given mask. 
	bds_dsmCmn_errListSize_DU8: USINT := 32;
	///Buffer size of error List (DTCs/DFCs) for a given mask
	bds_dsmCmn_dfesSize_DU8: USINT := 32;
END_VAR

// I/O API/IN legacy/GVL/GVL_in
VAR_GLOBAL
	///initialization after startup
	initIn_DB16: USINT := 16#1;
	///configured for AIV thresholds 
	cfgAiv_DB16: USINT := 16#2;
	///configured for AIC thresholds
	cfgAic_DB16: USINT := 16#4;
	///configured for AID thresholds 
	cfgAid_DB16: USINT := 16#8;
	///configured for RI thresholds
	cfgRi_DB16: USINT := 16#10;
	///configured for standard frequency sensor 
	cfgFreq_DB16: USINT := 16#20;
	///configured for DSM frequency sensor
	cfgFreqDSM_DB16: USINT := 16#40;
	lostSignalInfoDSM_DB16: USINT := 16#80;
	///shunt is activated for DSM sensor respective AIC
	actShunt_DB16: UINT := 16#1000;
	///locked shunt reactivation 
	lockReactShunt_DB16: UINT := 16#2000;
	cfgInMask_DB16: UINT := (((((cfgFreqDSM_DB16 OR cfgFreq_DB16) OR cfgRi_DB16) OR cfgAid_DB16) OR cfgAic_DB16) OR cfgAiv_DB16);
	///standstill
	standstill_DU8: USINT := 16#0;
	///direction left 
	dirLeft_DU8: USINT := 16#1;
	///direction right 
	dirRight_DU8: USINT := 16#2;
	///direction not known for sure (e.g. after standstill)
	dirUnknown_DU8: USINT := 16#4;
	/// error free 
	noError_DU8: USINT := 16#0;
	///air gap error (pulse is shorter than 64us)
	airGapError_DU8: USINT := 16#1;
	///mounting error (pulse is longer than 254us) 
	mountError_DU8: USINT := 16#2;
	///undefined signal length - should not occur (pulse is longer than 1785us
	signalLengthError_DU8: USINT := 16#4;
	///period too long or measured period exceeds maximum period 
	signalError_DU8: USINT := 16#8;
	///no status signal available (frequency to high)
	noStatusAvailable_DU8: USINT := 16#10;
	diagSCUBAT_DU8: USINT := 16#20;
	diagSCGND_OR_OL_DU8: USINT := 16#40;
	///DSM mask to get the frequency out
	maskFrequency_DU32: UDINT := 16#FFFFF;
	///DSM mask to get the direction
	maskDirection_DU32: UDINT := 16#F00000;
	///DSM shift number to get the direction
	numShiftDirection_DU32: USINT := 20;
	///DSM mask to get the status
	maskStatus_DU32: UDINT := 16#FF000000;
	///DSM shift number to get the status
	numShiftStatus_DU32: USINT := 24;
	///no period measured for phase signal 1
	lostPhaseSignal_1_DU8: USINT := 16#1;
	///no period measured for phase signal 2
	lostPhaseSignal_2_DU8: USINT := 16#2;
	SENT_STATUS_DRIVER_INIT_DU32: USINT := 16#1;
	SENT_STATUS_DRIVER_RUNNING_DU32: USINT := 16#2;
	SENT_STATUS_ONE_FRAME_RECEIVED_DU32: USINT := 16#4;
	SENT_STATUS_NEW_FRAME_RECEIVED_DU32: USINT := 16#8;
	SENT_STATUS_ONE_SLOW_FRAME_RECEIVED_DU32: USINT := 16#10;
	SENT_STATUS_NEW_SLOW_FRAME_RECEIVED_DU32: USINT := 16#20;
	SENT_ERROR_LINE_LOW_DU32: USINT := 16#40;
	SENT_ERROR_LINE_HIGH_DU32: USINT := 16#80;
	SENT_ERROR_NODAT_DU32: UINT := 16#100;
	SENT_ERROR_NOSIG_DU32: UINT := 16#200;
	SENT_ERROR_NOISE_DU32: UINT := 16#400;
	SENT_ERROR_DEBOUNCING_DU32: UINT := 16#800;
	SENT_ERROR_CRC_DU32: UINT := 16#1000;
	SENT_ERROR_RANGE_DU32: UINT := 16#2000;
	SENT_ERROR_MISSING_NIBBLE_DU32: UINT := 16#4000;
	SENT_ERROR_TOOMANY_NIBBLES_DU32: UINT := 16#8000;
	SENT_ERROR_MSG_LOST_DU32: UDINT := 16#10000;
	SENT_ERROR_SLOW_CRC_DU32: UDINT := 16#20000;
	SENT_ERROR_SLOW_MISSING_FRAME_DU32: UDINT := 16#40000;
	SENT_ERROR_NOSLOWDAT_DU32: UDINT := 16#80000;
	SENT_ERROR_CAL_PULSE_RANGE_DU32: UDINT := 16#100000;
	SENT_ERROR_CAL_SUCCESSIVE_DEVIATION_DU32: UDINT := 16#200000;
	SENT_WARNING_CAL_DEVIATION_20PCT_DU32: UDINT := 16#400000;
	SENT_ERROR_PAUSE_PULSE_RANGE_DU32: UDINT := 16#800000;
	SENT_ERROR_FAST_DATA_CTR_DU32: UDINT := 16#1000000;
	SENT_ERROR_FAST_DATA_INV_MSN0_DU32: UDINT := 16#2000000;
	NTC: USINT := 16#11;
	PTC: USINT := 16#22;
END_VAR

// Communication API/ISOBUS/GVL/GVL_isobus
VAR_GLOBAL
	///isobus rx/tx databox status
	BDS_ISOBUS_BOXSTATUS_NONE_DU16: UINT := 16#0;
	///isobus rx/tx databox status
	BDS_ISOBUS_BOXSTATUS_INIT_DU16: UINT := 16#100;
	///isobus rx/tx databox status
	BDS_ISOBUS_BOXSTATUS_VALID_DU16: UINT := 16#200;
	///isobus rx/tx databox status
	BDS_ISOBUS_BOXSTATUS_VAL_OVFL_DU16: UINT := 16#201;
	///isobus rx/tx databox status
	BDS_ISOBUS_BOXSTATUS_INV_SEQNBR_DU16: UINT := 16#301;
	///isobus rx/tx databox status
	BDS_ISOBUS_BOXSTATUS_INV_ABORT_DU16: UINT := 16#302;
	///isobus rx/tx databox status
	BDS_ISOBUS_BOXSTATUS_INV_TIMEOUT_DU16: UINT := 16#303;
	///isobus rx/tx databox status
	BDS_ISOBUS_BOXSTATUS_INV_OVFL_DU16: UINT := 16#304;
	///isobus rx/tx databox status
	BDS_ISOBUS_BOXSTATUS_INV_PGN_ERR_DU16: UINT := 16#310;
	///isobus rx/tx databox status
	BDS_ISOBUS_BOXSTATUS_INV_DPO_ERR_DU16: UINT := 16#311;
	///isobus rx/tx databox status
	BDS_ISOBUS_BOXSTATUS_PENDING_DU16: UINT := 16#400;
	///isobus rx/tx databox status
	BDS_ISOBUS_BOXSTATUS_BAM_RX_DU16: UINT := 16#500;
	///isobus rx/tx databox status
	BDS_ISOBUS_BOXSTATUS_CMDT_RX_DU16: UINT := 16#501;
	///isobus rx/tx databox status
	BDS_ISOBUS_BOXSTATUS_BAM_TX_DU16: UINT := 16#600;
	///isobus rx/tx databox status
	BDS_ISOBUS_BOXSTATUS_UNPACK_DU16: UINT := 16#700;
	///isobus rx/tx databox status
	BDS_ISOBUS_BOXSTATUS_ETP_RX_DU16: UINT := 16#800;
	///isobus rx/tx databox status
	BDS_ISOBUS_BOXSTATUS_MASK_DU16: UINT := 16#FF00;
	///isobus controller application status  (main status = hi byte, sub status = lo byte)
	BDS_ISOBUS_CASTATUS_NONE_DU16: UINT := 16#0;
	///isobus controller application status  (main status = hi byte, sub status = lo byte)
	BDS_ISOBUS_CASTATUS_INIT_DU16: UINT := 16#100;
	///isobus controller application status  (main status = hi byte, sub status = lo byte)
	BDS_ISOBUS_CASTATUS_WAIT_CLAIM_DU16: UINT := 16#200;
	///isobus controller application status  (main status = hi byte, sub status = lo byte)
	BDS_ISOBUS_CASTATUS_ADDR_CLAIMED_DU16: UINT := 16#300;
	///isobus controller application status  (main status = hi byte, sub status = lo byte)
	BDS_ISOBUS_CASTATUS_CANNOT_CLAIM_DU16: UINT := 16#400;
	///isobus controller application status  (main status = hi byte, sub status = lo byte)
	BDS_ISOBUS_CASTATUS_MASK_DU16: UINT := 16#FF00;
	///This sub status is automatically reset after a request via API function |bds_isobus_getStatus|
	BDS_ISOBUS_SUBSTATUS_TIMEOUT_DU16: UINT := 16#1;
	///This sub status is automatically reset after a request via API function |bds_isobus_getStatus|
	BDS_ISOBUS_SUBSTATUS_RXOVFL_DU16: UINT := 16#2;
	///This sub status is automatically reset after a request via API function |bds_isobus_getStatus|
	BDS_ISOBUS_SUBSTATUS_RESET_MASK_DU16: UINT := 16#FFF0;
	///This sub status is automatically reset after a request via API function |bds_isobus_getStatus|
	BDS_ISOBUS_SUBSTATUS_STOP_BC_DM13_DU16: UINT := 16#10;
	BDS_ISOBUS_RC_NO_ERRORS_DU16: UINT := 0;
	BDS_ISOBUS_RC_INVALID_ADDR_DU16: UINT := 1;
	BDS_ISOBUS_RC_INV_DATABOX_DU16: UINT := 2;
	BDS_ISOBUS_RC_INV_PGN_DU16: UINT := 3;
	BDS_ISOBUS_RC_INV_SRC_DU16: UINT := 4;
	BDS_ISOBUS_RC_INV_TIMEOUT_DU16: UINT := 5;
	BDS_ISOBUS_RC_INV_DATA_LEN_DU16: UINT := 6;
	BDS_ISOBUS_RC_INV_DATA_PTR_DU16: UINT := 7;
	BDS_ISOBUS_RC_OVERLAP_ADDR_DU16: UINT := 8;
	BDS_ISOBUS_RC_INV_STARTTIMEOUT_DU16: UINT := 9;
	BDS_ISOBUS_RC_INV_CYCLE_DU16: UINT := 10;
	BDS_ISOBUS_RC_INV_OFFSET_DU16: UINT := 11;
	BDS_ISOBUS_RC_INV_PRIO_DU16: UINT := 12;
	BDS_ISOBUS_RC_PGN_SRC_EXIST_DU16: UINT := 20;
	BDS_ISOBUS_RC_PGN_PRIO_EXIST_DU16: UINT := 21;
	BDS_ISOBUS_RC_CFG_NOTALLOWED_DU16: UINT := 22;
	BDS_ISOBUS_RC_INV_BOX_STATUS_DU16: UINT := 30;
	BDS_ISOBUS_RC_INV_SPN_DU16: UINT := 40;
	BDS_ISOBUS_RC_INV_FMI_DU16: UINT := 41;
	BDS_ISOBUS_RC_DM1_FULL_DU16: UINT := 42;
	BDS_ISOBUS_RC_DM2_FULL_DU16: UINT := 43;
	BDS_ISOBUS_RC_SPN_NOT_FOUND_DU16: UINT := 44;
	BDS_ISOBUS_RC_INV_ECU_ADDR_DU16: UINT := 50;
	BDS_ISOBUS_RC_INV_DM_TYPE_DU16: UINT := 51;
	BDS_ISOBUS_RC_INV_LIST_SIZE_DU16: UINT := 60;
	BDS_ISOBUS_RC_INV_EE_PAGE_DU16: UINT := 61;
	BDS_ISOBUS_RC_INV_EE_IDX_DU16: UINT := 62;
	BDS_ISOBUS_RC_INIT_MISSING_DU16: UINT := 63;
	BDS_ISOBUS_RC_EE_OVERLAPPING_DU16: UINT := 64;
	BDS_ISOBUS_RC_EEP_OVERFLOW_DU16: UINT := 70;
	BDS_ISOBUS_RC_INV_INST_NUM_DU16: UINT := 80;
	BDS_ISOBUS_RC_INV_CAN_CHNL_DU16: UINT := 81;
	BDS_ISOBUS_RC_INV_CA_ADDR_DU16: UINT := 82;
	BDS_ISOBUS_RC_CA_ADDR_IN_USE_DU16: UINT := 83;
	BDS_ISOBUS_RC_REGINST_NOT_ALLOWED_DU16: UINT := 84;
	BDS_ISOBUS_RC_INV_FUNC_SEQU_DU16: UINT := 85;
	BDS_ISOBUS_RC_PGN_USED_INTERNAL_DU16: UINT := 86;
	BDS_ISOBUS_RC_DM1_NOT_EXIST_DU16: UINT := 0;
	BDS_ISOBUS_RC_DM1_EXIST_DU16: UINT := 1;
	BDS_ISOBUS_SPN_ALL_DU32: UDINT := 16#FFFFFFFF;
	BDS_ISOBUS_FMI_ALL_DU8: USINT := 16#FF;
	BDS_ISOBUS_BYTES_ALL_DU32: UDINT := 16#FFFFFFFF;
	BDS_ISOBUS_OWN_SN_DU32: UDINT := 16#FFFFFFFF;
	BDS_ISOBUS_LIST_NONE_DU16: UINT := 16#0;
	BDS_ISOBUS_LIST_DM1_DU16: UINT := 16#1;
	BDS_ISOBUS_LIST_DM2_DU16: UINT := 16#2;
	BDS_ISOBUS_LIST_DM1_V1_DU16: UINT := 16#11;
	BDS_ISOBUS_LIST_DM2_V1_DU16: UINT := 16#12;
	BDS_ISOBUS_LIST_DM1_V2_DU16: UINT := 16#21;
	BDS_ISOBUS_LIST_DM2_V2_DU16: UINT := 16#22;
	BDS_ISOBUS_LIST_DM1_V3_DU16: UINT := 16#31;
	BDS_ISOBUS_LIST_DM2_V3_DU16: UINT := 16#32;
	BDS_ISOBUS_DTC_LIST_SIZE_DU16: UINT := 20;
	///Maximum number of own DTCs within DTC list
	BDS_ISOBUS_MaxNbrDtc_DU16: UINT := 32;
	///Max data length of the ReqPgn TX databox buffer, the data of all requested PGNs(except the PGNs of the application TX-Boxes) must fit into this buffer!
	BDS_ISOBUS_buffLenReqPgn_DU16: UINT := 300;
	///Maximum size of a single message
	BDS_ISOBUS_MaxSingleSize_DU32: UDINT := 8;
	///Maximum size of a BAM/CMDT message
	BDS_ISOBUS_MaxTpSize_DU32: UDINT := 1785;
	///Maximum size of a ETP message
	BDS_ISOBUS_MaxETpSize_DU32: UDINT := 117440512;
	///Max data length of a DM1/2 TX databox buffer
	BDS_ISOBUS_DmBuffSize_DU16: UINT := 130;
	BDS_ISOBUS_QUEUE_OVERFLOW_DU8: USINT := 1;
	BDS_ISOBUS_QUEUE_UPDATED_DU8: USINT := 2;
	BDS_ISOBUS_QUEUE_UNDERFLOW_DU8: USINT := 3;
	BDS_ISOBUS_QUEUE_ELEMENT_DELETED_DU8: USINT := 4;
END_VAR

// Communication API/LIN/GVL/GVL_lin
VAR_GLOBAL
	BDS_LIN_ERR_NO_ERRORS_DU16: UINT := 0;
	BDS_LINSIG_ERR_NUM_TX_SIG_DU16: UINT := BDS_CANSIG_ERR_NUM_TX_SIG_DU16;
	BDS_LINSIG_ERR_NUM_RX_SIG_DU16: UINT := BDS_CANSIG_ERR_NUM_RX_SIG_DU16;
	BDS_LINSIG_ERR_TX_DATAPTR_DU16: UINT := BDS_CANSIG_ERR_TX_DATAPTR_DU16;
	BDS_LINSIG_ERR_RX_DATAPTR_DU16: UINT := BDS_CANSIG_ERR_RX_DATAPTR_DU16;
	BDS_LINSIG_ERR_TX_FAIL_DU16: UINT := BDS_CANSIG_ERR_TX_FAIL_DU16;
	BDS_LINSIG_ERR_RX_FAIL_DU16: UINT := BDS_CANSIG_ERR_RX_FAIL_DU16;
	BDS_LINSIG_ERR_TX_NOSERVICE_DU16: UINT := BDS_CANSIG_ERR_TX_NOSERVICE_DU16;
	BDS_LINSIG_ERR_RX_NOSERVICE_DU16: UINT := BDS_CANSIG_ERR_RX_NOSERVICE_DU16;
	BDS_LINSIG_ERR_RX_LENPTR_DU16: UINT := BDS_CANSIG_ERR_RX_LENPTR_DU16;
	BDS_LIN_INVALID_CHNL_DU16: UINT := 121;
	BDS_LIN_INVALID_SCHTABLE_NO_DU16: UINT := 122;
	BDS_LIN_ERR_NULLPOINTER_DU16: UINT := 123;
	BDS_LIN_TX_OK_DU8: USINT := 1;
	BDS_LIN_TX_BUSY_DU8: USINT := 2;
	BDS_LIN_TX_HEADER_ERROR_DU8: USINT := 3;
	BDS_LIN_TX_ERROR_DU8: USINT := 4;
	BDS_LIN_RX_OK_DU8: USINT := 5;
	BDS_LIN_RX_BUSY_DU8: USINT := 6;
	BDS_LIN_RX_ERROR_DU8: USINT := 7;
	BDS_LIN_RX_NO_RESPONSE_DU8: USINT := 8;
	BDS_LIN_OPERATIONAL_DU8: USINT := 9;
	BDS_LIN_CH_SLEEP_DU8: USINT := 10;
END_VAR

// Memory API/NVM/GVL/GVL_mem
VAR_GLOBAL
	///NVM block types
	BDS_MEM_BLOCKTYPE_APPL_DU16: UINT := 0;
	///NVM block types
	BDS_MEM_BLOCKTYPE_SYSTEM_DU16: UINT := 1;
	///function return codes
	BDS_MEM_NO_ERROR_DU16: UINT := 16#0;
	///function return codes
	BDS_MEM_INVALID_BLOCKID_DU16: UINT := 16#1;
	///function return codes
	BDS_MEM_INVALID_ADDRESS_DU16: UINT := 16#2;
	///function return codes
	BDS_MEM_BLOCK_INIT_DU16: UINT := 16#10;
	///function return codes
	BDS_MEM_READBLOCK_ERROR_DU16: UINT := 16#100;
	///function return codes
	BDS_MEM_WRITEBLOCK_ERROR_DU16: UINT := 16#200;
	///function return codes
	BDS_MEM_MARKBLOCK_ERROR_DU16: UINT := 16#400;
	///function return codes
	BDS_MEM_READBLOCK_DATASIZE_INVALID_DU16: UINT := 16#300;
	///function return codes
	BDS_MEM_WRITEBLOCK_DATASIZE_INVALID_DU16: UINT := 16#300;
	///function return codes
	BDS_MEM_WRITEBLOCK_DATAPTR_INVALID_DU16: UINT := 16#301;
	///function return codes
	BDS_MEM_READBLOCK_DATAPTR_INVALID_DU16: UINT := 16#301;
	///function return codes
	BDS_MEM_FFI_ACCESS_ERROR_DU16: UINT := 12;
	BDS_MEM_GETBLOCKSTATUS_ERROR_DU16: UINT := 16#300;
	BDS_MEM_REQ_FAILED_DU16: UINT := 16#301;
	BDS_MEM_REQ_PENDING_DU16: UINT := 16#302;
	BDS_MEM_REQ_INTEGRITY_FAILED_DU16: UINT := 16#303;
	BDS_MEM_REQ_BLOCK_SKIPPED_DU16: UINT := 16#304;
	BDS_MEM_REQ_NV_INVALIDATED_DU16: UINT := 16#305;
	BDS_MEM_REQ_CANCELED_DU16: UINT := 16#306;
	BDS_MEM_REQ_REDUNDANCY_FAILED_DU16: UINT := 16#307;
	BDS_MEM_REQ_RESTORED_FROM_ROM_DU16: UINT := 16#308;
	bds_mem_nvmBlock01_512_R_D: UINT := 13;
	bds_mem_nvmBlock02_512_R_D: UINT := 33;
	bds_mem_nvmBlock03_512_R_D: UINT := 47;
	bds_mem_nvmBlock04_512_R_D: UINT := 58;
	bds_mem_nvmBlock05_256_R_D: UINT := 15;
	bds_mem_nvmBlock06_256_R_D: UINT := 35;
	bds_mem_nvmBlock07_256_R_D: UINT := 49;
	bds_mem_nvmBlock08_256_R_D: UINT := 60;
	bds_mem_nvmBlock09_256_R_D: UINT := 17;
	bds_mem_nvmBlock10_256_R_D: UINT := 37;
	bds_mem_nvmBlock11_256_R_D: UINT := 51;
	bds_mem_nvmBlock12_256_R_D: UINT := 62;
	bds_mem_nvmBlock13_128_R_D: UINT := 20;
	bds_mem_nvmBlock14_128_R_D: UINT := 40;
	bds_mem_nvmBlock15_128_R_D: UINT := 54;
	bds_mem_nvmBlock16_128_R_D: UINT := 65;
	bds_mem_nvmBlock17_32_R_D: UINT := 23;
	bds_mem_nvmBlock18_32_R_D: UINT := 43;
	bds_mem_nvmBlock19_512_N_D: UINT := 12;
	bds_mem_nvmBlock20_512_N_D: UINT := 32;
	bds_mem_nvmBlock21_512_N_D: UINT := 46;
	bds_mem_nvmBlock22_512_N_D: UINT := 57;
	bds_mem_nvmBlock23_256_N_D: UINT := 14;
	bds_mem_nvmBlock24_256_N_D: UINT := 34;
	bds_mem_nvmBlock25_256_N_D: UINT := 48;
	bds_mem_nvmBlock26_256_N_D: UINT := 59;
	bds_mem_nvmBlock27_256_N_D: UINT := 16;
	bds_mem_nvmBlock28_256_N_D: UINT := 36;
	bds_mem_nvmBlock29_256_N_D: UINT := 50;
	bds_mem_nvmBlock30_256_N_D: UINT := 61;
	bds_mem_nvmBlock31_128_N_D: UINT := 19;
	bds_mem_nvmBlock32_128_N_D: UINT := 39;
	bds_mem_nvmBlock33_128_N_D: UINT := 53;
	bds_mem_nvmBlock34_128_N_D: UINT := 64;
	bds_mem_nvmBlock35_32_N_D: UINT := 22;
	bds_mem_nvmBlock36_32_N_D: UINT := 42;
	bds_mem_nvmBlock37_64_N_D: UINT := 24;
	bds_mem_nvmBlock38_64_N_D: UINT := 44;
	bds_mem_nvmBlock39_64_N_D: UINT := 56;
	bds_mem_nvmBlock40_64_N_D: UINT := 67;
	bds_mem_nvmBlock41_64_N_D: UINT := 71;
	bds_mem_nvmBlock42_64_N_D: UINT := 75;
	bds_mem_nvmBlock43_64_N_D: UINT := 79;
	bds_mem_nvmBlock44_64_N_D: UINT := 82;
	bds_mem_nvmBlock45_64_N_D: UINT := 85;
	bds_mem_nvmBlock46_64_N_D: UINT := 88;
	bds_mem_nvmBlock47_128_R_D: UINT := 21;
	bds_mem_nvmBlock48_128_R_D: UINT := 41;
	bds_mem_nvmBlock49_128_R_D: UINT := 55;
	bds_mem_nvmBlock50_128_R_D: UINT := 66;
	bds_mem_nvmBlock51_128_R_D: UINT := 70;
	bds_mem_nvmBlock52_128_R_D: UINT := 74;
	bds_mem_nvmBlock53_128_R_D: UINT := 78;
	bds_mem_nvmBlock54_128_R_D: UINT := 81;
	bds_mem_nvmBlock55_128_R_D: UINT := 84;
	bds_mem_nvmBlock56_128_R_D: UINT := 87;
	bds_mem_nvmBlock57_128_R_D: UINT := 25;
	bds_mem_nvmBlock58_128_R_D: UINT := 26;
	bds_mem_nvmBlock59_128_R_D: UINT := 27;
	bds_mem_nvmBlock60_128_R_D: UINT := 28;
	bds_mem_nvmBlock61_128_R_D: UINT := 29;
	bds_mem_nvmBlock62_128_R_D: UINT := 30;
	bds_mem_nvmBlock63_256_R_D: UINT := 18;
	bds_mem_nvmBlock64_256_R_D: UINT := 38;
	bds_mem_nvmBlock65_256_R_D: UINT := 52;
	bds_mem_nvmBlock66_256_R_D: UINT := 63;
	bds_mem_nvmBlock67_256_R_D: UINT := 69;
	bds_mem_nvmBlock68_256_R_D: UINT := 73;
	bds_mem_nvmBlock69_256_R_D: UINT := 77;
	bds_mem_nvmBlock70_512_R_D: UINT := 68;
	bds_mem_nvmBlock71_512_R_D: UINT := 72;
	bds_mem_nvmBlock72_512_R_D: UINT := 76;
	bds_mem_nvmBlock73_512_R_D: UINT := 80;
	bds_mem_nvmBlock74_512_R_D: UINT := 83;
	bds_mem_nvmBlock75_512_R_D: UINT := 86;
	bds_mem_nvmBlock76_512_N_D: UINT := 11;
	bds_mem_nvmBlock77_1024_N_D: UINT := 10;
	bds_mem_nvmBlock78_1024_N_D: UINT := 31;
	bds_mem_nvmBlock79_1024_N_D: UINT := 45;
	BDS_MEM_INVALID_TABLE_MAPPING_DU16: UINT := 16#3;
	BDS_MEM_NVM_CANCONFIG_BLOCK_DU16: UINT := 113;
	BDS_MEM_BAUD_SMPLRATE_ADDR_DU8: USINT := 42;
	BDS_MEM_UDS_NODE_ID_ADDR_DU8: USINT := 43;
	BDS_MEM_UDS_TESTER_ID_ADDR_DU8: USINT := 44;
	BDS_MEM_UDS_RXTX_ID_LSB_ADDR_DU8: USINT := 45;
	BDS_MEM_UDS_RXTX_ID_MSB_ADDR_DU8: USINT := 46;
	BDS_MEM_UDS_ECONFIG_NODEID_DU8: USINT := 47;
	BDS_MEM_PBS_VRNT_ADDR_DU8: USINT := 63;
	BDS_MEM_CONFIG_INIT_DU8: USINT := 1;
	BDS_MEM_CONFIG_DEFAULT_DU8: USINT := 2;
	BDS_MEM_MPG_TABLE_ROW_DU8: USINT := 8;
	BDS_MEM_MPG_TABLE_COL_DU8: USINT := 2;
	BDS_MEM_MOVE_UPPER_NIBBLE_DU8: USINT := 4;
	BDS_MEM_DFT_CAN_CHANNEL_DU8: USINT := 2;
	BDS_MEM_DFT_CAN_BAUDRATE_DU32: UDINT := 250000;
	BDS_MEM_DFT_CAN_SAMPLING_POINT_DU8: USINT := 80;
	BDS_MEM_DFT_UDS_NODEID_DU8: USINT := 16#1;
	BDS_MEM_DFT_UDS_TESTERID_DU8: USINT := 16#FA;
	BDS_MEM_DFT_UDS_RXTXIDENTIFIERS_DU16: UINT := 16#18DA;
END_VAR

// I/O API/OUT/GVL/GVL_out
VAR_GLOBAL
	/// possible dither frequency value 
	fDither_0Hz_DU8: USINT := 0;
	/// possible dither frequency values 
	fDither_83Hz_DU8: USINT := 83;
	/// possible dither frequency values 
	fDither_90Hz_DU8: USINT := 90;
	/// possible dither frequency values 
	fDither_100Hz_DU8: USINT := 100;
	/// possible dither frequency values 
	fDither_111Hz_DU8: USINT := 111;
	/// possible dither frequency values 
	fDither_125Hz_DU8: USINT := 125;
	/// possible dither frequency values 
	fDither_142Hz_DU8: USINT := 142;
	/// possible dither frequency values 
	fDither_166Hz_DU8: USINT := 166;
	/// possible dither frequency values 
	fDither_200Hz_DU8: USINT := 200;
	/// possible dither frequency values 
	fDither_250Hz_DU8: USINT := 250;
	/// initialization after startup 
	initOut_DB16: USINT := 16#1;
	/// configuration of closed loop control 
	cfgPOC_DB16: USINT := 16#2;
	/// configuration of period 
	cfgPeriod_DB16: USINT := 16#4;
	/// configuration of dither 
	cfgDither_DB16: USINT := 16#8;
	/// configuration of deviation 
	cfgDeviation_DB16: USINT := 16#10;
	/// configuration of KpKi 
	cfgPI_DB16: USINT := 16#20;
	/// locked by SCB...necessary for AOV 
	lockedSCB_DB16: USINT := 16#40;
	/// locked by SCG...necessary for AOV 
	lockedSCG_DB16: USINT := 16#80;
	/// locked by OC 
	lockedOC_DB16: UINT := 16#100;
	/// locked by Error Handler 
	locked_DB16: UINT := 16#200;
	/// locked by Monitoring Module (MO) Error
	lockedMO_DB16: UINT := 16#400;
	/// locked reactivation timer reload after a hot short circuit 
	lockCouTiReact_DB16: UINT := 16#800;
	/// time for reactivation after a hot short circuit not elapsed 
	tiReactNotElapsed_DB16: UINT := 16#1000;
	/// linked at least with one other safout output 
	linked_DB16: UINT := 16#2000;
	/// Test pulses disable 
	tlsPlsDis_DB16: UINT := 16#4000;
	/// output is disabled (avoid open load faults of unused outputs)
	disabled_DB16: UINT := 16#8000;
	cfgOutMask_DB16: UINT := ((((cfgPI_DB16 OR cfgDeviation_DB16) OR cfgDither_DB16) OR cfgPeriod_DB16) OR cfgPOC_DB16);
	lockedMaskAOV_DB16: UINT := (lockedSCG_DB16 OR lockedSCB_DB16);
	lockedMaskFSC_DB16: UINT := ((lockedMO_DB16 OR locked_DB16) OR lockedOC_DB16);
	BDS_OUT_UNLOCK_OK_DU16: UINT := 16#0;
	BDS_OUT_UNLOCK_ERR_MO_DU16: UINT := 16#1;
	BDS_OUT_UNLOCK_ERR_REACT_CNT_DU16: UINT := 16#2;
	BDS_OUT_UNLOCK_ERR_SCB_DU16: UINT := 16#4;
	BDS_OUT_UNLOCK_ERR_SCG_DU16: UINT := 16#8;
	BDS_OUT_UNLOCK_ERR_OL_DU16: UINT := 16#10;
	BDS_OUT_UNLOCK_ERR_OT_DU16: UINT := 16#20;
	BDS_OUT_UNLOCK_ERR_OR_DU16: UINT := 16#40;
	BDS_OUT_UNLOCK_RES_OC_DU16: UINT := 16#80;
	BDS_OUT_UNLOCK_ERR_SIG_DU16: UINT := 16#8000;
END_VAR

// I/O API/SAFOUT/GVL/GVL_safout
VAR_GLOBAL
	/// initialization after startup 
	initialized_DB16: UDINT := 16#1;
	/// configured channel 
	configured_DB16: UDINT := 16#2;
	/// activated outputs 
	activeOut1_DB16: UDINT := 16#10;
	/// activated outputs 
	activeOut2_DB16: UDINT := 16#20;
	/// activated outputs 
	activeOut3_DB16: UDINT := 16#40;
	/// activated outputs 
	activeOut4_DB16: UDINT := 16#80;
	/// locked channel 
	lockedChnl_DB16: UDINT := 16#100;
	/// only for internal use 
	checkOut1_DB16: UDINT := 16#200;
	/// only for internal use 
	checkOut2_DB16: UDINT := 16#400;
	/// only for internal use 
	displayErrorHS_DB16: UDINT := 16#1000;
	/// maximal current deviation of the HS/LS compare is exceeded 
	iDevCmpHSLS_DB16: UDINT := 16#2000;
	/// ignore non critical faults 
	ignoreError_DB16: UDINT := 16#8000;
	activeOut_Mask_DB16: UDINT := 16#F0;
	/// number of channels 
	SAFOUT_CHNL_NUM_DU16: UINT := 5;
	/// Proportional Highside Digital lowside switchable safout mode 
	PHDLS: UDINT := 16#1100;
	/// Digital Highside Digital Lowside Multiple safout mode 
	DHDLM: UDINT := 16#2200;
	/// Proportional Highside Multiple Digital Lowside safout mode 
	PHMDL: UDINT := 16#3300;
	/// Proportional Lowside Digital Highside switchable safout mode 
	PLDHS: UDINT := 16#4400;
	/// Digital Lowside Digital Highside Multiple safout mode
	DLDHM: UDINT := 16#5500;
	/// Proportional Lowside Multiple Digital Highside safout mode
	PLMDH: UDINT := 16#6600;
	/// channel number 
	CHNL1: UDINT := 16#0;
	/// channel number 
	CHNL2: UDINT := 16#1;
	/// channel number 
	CHNL3: UDINT := 16#2;
	/// channel number 
	CHNL4: UDINT := 16#3;
	/// channel number 
	CHNL5: UDINT := 16#4;
	/// channel number 
	CHNL6: UDINT := 16#5;
	/// channel number 
	CHNL7: UDINT := 16#6;
	/// channel number 
	CHNL8: UDINT := 16#7;
	/// channel number 
	CHNL9: UDINT := 16#8;
	/// channel number 
	CHNL10: UDINT := 16#9;
	/// channel number 
	CHNL11: UDINT := 16#A;
	/// channel number 
	CHNL12: UDINT := 16#B;
	/// channel number 
	CHNL13: UDINT := 16#C;
	/// channel number 
	CHNL14: UDINT := 16#D;
	/// channel number 
	CHNL15: UDINT := 16#E;
	/// channel number 
	CHNL16: UDINT := 16#F;
	/// channel number 
	CHNL17: UDINT := 16#10;
	/// channel number 
	CHNL18: UDINT := 16#11;
	MASK_CHNL_DU16: UINT := 16#FF;
	MASK_MODE_DU16: UINT := 16#FF00;
	MASK_SIGNAL_DU16: UINT := 16#FF;
	MASK_SIGNAL_TYPE_DU16: UINT := 16#FF00;
	SIGNAL_TYPE_DO_DU16: UINT := (16#100 AND MASK_SIGNAL_TYPE_DU16);
	SIGNAL_TYPE_PO_DU16: UINT := (16#200 AND MASK_SIGNAL_TYPE_DU16);
	/// fault ordering (per nibble) of the diagnostic info 
	SAFOUT_SCB: UDINT := 16#1;
	/// fault ordering (per nibble) of the diagnostic info 
	SAFOUT_SCG: UDINT := 16#2;
	/// fault ordering (per nibble) of the diagnostic info 
	SAFOUT_OL: UDINT := 16#4;
	/// fault ordering (per nibble) of the diagnostic info 
	SAFOUT_OC: UDINT := 16#8;
	/// Safout test is enabled 
	safoutTestCfg_DU16: UINT := 16#1;
	/// Safout test is running 
	safoutTestAct_DU16: UINT := 16#2;
	/// Safout test is complete 
	safoutTestCmp_DU16: UINT := 16#4;
END_VAR

// System API/SEC/GVL/GVL_sec
VAR_GLOBAL
	///default security level
	BDS_SEC_DEFAULT_SEC_LEVEL_DU8: USINT := 0;
	BDS_SEC_MIN_ASW_SEC_LEVEL_DU8: USINT := 1;
	BDS_SEC_MAX_ASW_SEC_LEVEL_DU8: USINT := 10;
	///min. random number length in bds_sec_getRnd
	BDS_SEC_MIN_RANDOM_LENGTH_DU16: UINT := 1;
	///max. random number length in bds_sec_getRnd
	BDS_SEC_MAX_RANDOM_LENGTH_DU16: UINT := 512;
	BDS_SEC_ERR_NO_ERROR_DU16: UINT := 16#0;
	BDS_SEC_ERR_PARAM1_ERROR_DU16: UINT := 16#1;
	BDS_SEC_ERR_PARAM2_ERROR_DU16: UINT := 16#2;
	BDS_SEC_ERR_PARAM3_ERROR_DU16: UINT := 16#3;
	BDS_SEC_ERR_PARAM4_ERROR_DU16: UINT := 16#4;
	BDS_SEC_ERR_REQUEST_PENDING_DU16: UINT := 16#10;
	BDS_SEC_ERR_WAIT_FOR_STARTUP_DELAY_DU16: UINT := 16#11;
	BDS_SEC_ERR_INVALID_SEQUENCE_DU16: UINT := 16#20;
	BDS_SEC_ERR_NBR_ATTEMPTS_EXCEEDED_DU16: UINT := 16#21;
	BDS_SEC_ERR_HSM_NOT_ACTIVE_DU16: UINT := 16#30;
	BDS_SEC_ERR_INITIALIZATION_FAILED_DU16: UINT := 16#31;
	BDS_SEC_ERR_GET_SEED_FAILED_DU16: UINT := 16#32;
	BDS_SEC_ERR_OPEN_SESSION_FAILED_DU16: UINT := 16#33;
	BDS_SEC_ERR_GENERATE_RANDOM_FAILED_DU16: UINT := 16#34;
	BDS_SEC_ERR_CLOSE_SESSION_FAILED_DU16: UINT := 16#35;
	BDS_SEC_ERR_ENCRYPT_INIT_FAILED_DU16: UINT := 16#36;
	BDS_SEC_ERR_ENCRYPT_FAILED_DU16: UINT := 16#37;
	BDS_SEC_ERR_SET_PASSWORD_FAILED_DU16: UINT := 16#38;
	BDS_SEC_ERR_COMPARE_KEY_Faild_DU16: UINT := 16#39;
	BDS_SEC_SECDATA_LENGTH_DU32: UDINT := 16;
END_VAR

// System API/SYS/GVL/GVL_sys
VAR_GLOBAL
	OperatingHour_updatefrequency_DU16: UINT := 1800;
	BDS_VERSION_SW_PART_APPL_DU8: USINT := 16#0;
	BDS_VERSION_SW_PART_SB_DU8: USINT := 16#1;
	BDS_VERSION_SW_PART_CB_DU8: USINT := 16#2;
	BDS_VERSION_SW_PART_BSW_NAME_DU8: USINT := 16#3;
	BDS_VERSION_SW_PART_BSW_VERSION_DU8: USINT := 16#4;
	BDS_VERSION_SW_PART_EC_PROJECT_DU8: USINT := 16#5;
	BDS_SYSGETVERSION_OK_DU16: UINT := 16#0;
	BDS_SYSGETVERSION_BUFLEN_UNDERSIZE_DU16: UINT := 16#1;
	BDS_SYSGETVERSION_SW_PART_INVALID_DU16: UINT := 16#2;
	BDS_SYSGETVERSION_SW_INFO_NOT_FOUND_DU16: UINT := 16#3;
	BDS_SYSGETVERSION_BUF_INVALID_DU16: UINT := 16#4;
	BDS_SYSGETVERSION_COPIEDBYTES_INVALID_DU16: UINT := 16#5;
	BDS_SYS_DISABLE_PROLONG_PSTDRV_DL: UINT := 16#0;
	BDS_SYS_ENABLE_PROLONG_PSTDRV_DL: UINT := 16#1;
	BDS_MAX_NBR_ERR_CODES_DU16: UINT := 20;
	EEPPAGE_API_DU16: UINT := 15;
	EEPPAGE_APPL1_BEGIN_DU16: UINT := 1;
	EEPPAGE_APPL1_END_DU16: UINT := 14;
	EEPPAGE_APPL2_BEGIN_DU16: UINT := 32;
	EEPPAGE_APPL2_END_DU16: UINT := 60;
	BDS_SYS_ERR_SWNM_DU16: UINT := 1;
	BDS_SYS_ERR_HWID_DU16: UINT := 2;
	BDS_SYS_MAX_SWNM_LEN_DU16: UINT := 50;
	BDS_SYS_ERR_INVALID_API_DU16: UINT := 4;
	BDS_SYS_NO_ERROR_DU16: UINT := 0;
	BDS_SYS_PARAM1_ERROR_DU16: UINT := 1;
	BDS_SYS_PARAM2_ERROR_DU16: UINT := 2;
	BDS_SYS_FAULT_PERCENT_100_DU8: USINT := 15;
	E_NOT_OK: USINT := 16#1;
	E_OK: USINT := 16#0;
	STD_HIGH: USINT := 16#1;
	STD_LOW: USINT := 16#0;
	STD_ACTIVE: USINT := 16#1;
	STD_IDLE: USINT := 16#0;
	STD_ON: USINT := 16#1;
	STD_OFF: USINT := 16#0;
	BDS_WAKE_T15_DU32: UDINT := 16#15;
	BDS_WAKE_CAN4_DU32: UDINT := 16#4;
	BDS_WAKE_CAN1_DU32: UDINT := 16#1;
	BDS_SYS_OPERHRSREADTIMEINTERVAL_DU16: UINT := 1780;
	BDS_SYS_MAXOPERHRS_DU32: UDINT := 16#FFFFFFFE;
	BDS_SYS_ERR_PARA_INVALID_DU8: USINT := 2;
	BDS_SYS_ERR_INVALID_INPUT_DU8: USINT := 3;
	BDS_SYS_ERR_OPERHRS_DU32: UDINT := 16#1;
	BDS_SYS_FFI_ACCESS_ERROR_DU8: USINT := 25;
	BDS_SYS_FFI_ACCESS_ERROR_GETVALUE_DU32: UDINT := 0;
	BDS_SYS_FFI_ACCESS_ERROR_GETVALUE_DU64: ULINT := 0;
END_VAR

// Diagnostics API/UDS/GVL/GVL_uds
VAR_GLOBAL
	UDS_PREVENT_ALL_DU8: USINT := 16#0;
	UDS_PERMIT_ALL_DU8: USINT := 16#FF;
	UDS_ERR_NOT_CALLED_IN_SYS_DU8: USINT := 16#FF;
	UDS_SOFTRESET_ACCESS_DU8: USINT := 16#1;
	UDS_HARDRESET_ACCESS_DU8: USINT := 16#2;
	UDS_KEYOFFONRESET_ACCESS_DU8: USINT := 16#4;
	UDS_PROGRAMMINGSESS_ACCESS_DU8: USINT := 16#10;
	BDS_UDS_ERR_PARA_INVALID_DU8: USINT := 16#2;
	BDS_UDS_ERR_NODEID_DU8: USINT := 16#3;
	BDS_UDS_MASKING_BITS_DU16: UINT := 16#1FFF;
	BDS_UDS_FFI_ACCESS_ERROR_DU16: UINT := 25;
	BDS_UDS_NODEID_DU8: USINT := 16#1;
	BDS_UDS_TESTERID_DU8: USINT := 16#FA;
	BDS_UDS_RXTXIDENTIFIERS_DU16: UINT := 16#18DA;
	BDS_UDS_CAN_CHANNEL_DU8: USINT := 2;
	BDS_UDS_CAN_BAUDRATE_DU32: UDINT := 250000;
	BDS_UDS_CAN_SAMPLING_POINT_DU8: USINT := 80;
END_VAR

// Diagnostics API/XCP/GVL/GVL_xcp
VAR_GLOBAL
	///Disable XCP communication.
	BDS_DISABLE_XCP_DU16: UINT := 16#0;
	///Enable read, write Access in XCP.
	BDS_ENABLE_XCP_DU16: UINT := 16#FFFF;
	///Enable read only Access in XCP.
	BDS_ENABLE_XCP_READ_DU16: UINT := 16#FFFE;
END_VAR

// Communication API/CAN/CAN legacy/API/bds_can_getData
///Get the oldest message (FIFO) FROM the receive buffer OF the specified CAN channel.
///
///=======
/// Remarks:
///=======
///	+ A CAN receive buffer is NOT available UNTIL a buffer is registered within easyConfig.
///	+ Only received data with identifiers which does NOT match with identifiers OF initialized receive data boxes are saved AND can be read BY using THIS FUNCTION!
///    + First check the RETURN value before accessing the message.
///    + The |GVL_can| is given for usage of defines.
///----------
/// CAUTION:
///----------
///If the ISOBUS module is used then the CAN receive buffer on the corresponding CAN channel is exclusively used by ISOBUS. In this case this function must not be used any more by the application!
///
///----------
/// FFI:
///----------
///This API can be used in trusted partitions. For untrusted partitions use |bds_can_getData_ffi|. See Freedom from Interference (FFI) concept for more details.
///
///==================================================================		  			===================================================================================================
///Return value    								  									Description
///==================================================================		  			===================================================================================================
///0: BDS_CAN_ERR_NO_ERRORS_DU16					  									Function is called without errors. Message data returned in msg_s are valid.
///14: BDS_CAN_ERR_CHNL_DU16						  									Unknown CAN channel.
///30: BDS_CAN_ERR_RXBUF_OVFL_DU16					  									Receive buffer overflow. At least one message is lost. Message data returned in msg_s are valid.
///31: BDS_CAN_ERR_RXBUF_EMPTY_DU16				  										Receive buffer is empty. Message data returned in msg_s are invalid.
///32: BDS_CAN_ERR_RXBUF_LEN0_DU16														Receive buffer length is zero. Message data returned in msg_s are invalid.
///60: BDS_CAN_ERR_INVALID_ADDR_DU16													Invalid address (parameter msg_s).
///5: BDS_CAN_FFI_ACCESS_ERROR_DU16														FFI API access error.
///
///==================================================================		   			===================================================================================================
///
///=======
///Code Example:
///=======
///============================================================================
///
///PROGRAM appl_Task_1
///  VAR
///     msg_s: bds_can_Message_ts;
///  END_VAR
///
///  IF (0 = bds_can_getData(BDS_CAN_1_D, ADR(msg_s))) THEN
///  
///    (* Message in structure msg_s is valid and can be evaluated. *)
///	
///  END_IF
///END
///
///============================================================================
{attribute 'external_name' := 'cmp_rts_bds_can_getData'}
FUNCTION bds_can_getData : UINT
VAR_INPUT
	///Indicates the CAN channel.Possible values are
	///    + BDS_CAN_1_D(0)
	///    + BDS_CAN_2_D(1)
	///    + BDS_CAN_3_D(2)
	///	+ BDS_CAN_4_D(3)
	chnl_e: bds_can_Chnl_te;
	///Pointer to the message data of type bds_can_Message_ts.
	msg_ps: POINTER TO bds_can_Message_ts;
END_VAR

END_FUNCTION

// Communication API/CAN/CAN_FFI_API/bds_can_getData_ffi
{attribute 'external_name' := 'cmp_rts_bds_can_getData_ffi'}
FUNCTION bds_can_getData_ffi : UINT
VAR_INPUT
	///Indicates the CAN channel.Possible values are
	///    + BDS_CAN_1_D(0)
	///    + BDS_CAN_2_D(1)
	///    + BDS_CAN_3_D(2)
	///	+ BDS_CAN_4_D(3)
	chnl_e: bds_can_Chnl_te;
	///Pointer to the message data of type bds_can_Message_ts.
	msg_ps: POINTER TO bds_can_Message_ts;
END_VAR

END_FUNCTION

// Communication API/CAN/CAN legacy/API/bds_can_getDatabox
///Gets a message from the specified receive databox of the specified CAN channel.
///
///=======
/// Remarks:
///=======
///	+ The specified receive databox has to be initialized by |bds_can_initRxDatabox| before using this function.
///	+ If the databox was initialized with a buffer length = 1 then the last received message will be read from the databox buffer.
///	+ If the databox was initialized with a buffer length > 1 then the oldest message will be read from the databox buffer.
///	+ The number of required receive databoxes must be defined by easyConfig before using this function.
///    + The |GVL_can| is given for usage of defines.
///
///==================================================================		  			===================================================================================================
///Return value    								  									Description
///==================================================================		  			===================================================================================================
///0: BDS_CAN_ERR_NO_ERRORS_DU16					  									Function is called without errors. Message data returned in data_pau8 are valid.
///9: BDS_CAN_ERR_DATABOXNUM_DU16					  									Invalid databox number.
///14: BDS_CAN_ERR_CHNL_DU16					  										Unknown CAN channel.
///30: BDS_CAN_ERR_RXBUF_OVFL_DU16					  									Receive buffer overflow. At least one message is lost. Message data returned in msg_s are valid.
///31: BDS_CAN_ERR_RXBUF_EMPTY_DU16					  								Receive buffer is empty. Message data returned in msg_s are invalid.
///60: BDS_CAN_ERR_INVALID_ADDR_DU16					  								Invalid address (parameter msg_s).
///62: BDS_CAN_ERR_DATABOX_NOINIT_DU16					  								Databox is not initialized.
///5: BDS_CAN_FFI_ACCESS_ERROR_DU16														FFI API access error.
///==================================================================		   			===================================================================================================
///
///----------
/// FFI:
///----------
///This API can be used in trusted partitions only. For untrusted partitions use |bds_can_getDatabox_ffi|. See Freedom from Interference (FFI) concept for more details.
///
///=======
///Code Example:
///=======
///============================================================================
///
///PROGRAM can_1_RxDatabox_1_Callback
///  VAR
///    DataboxData_au8: ARRAY[1..8] of USINT;
///    DataboxNumBytes_u8: USINT;
///  END_VAR
///
///  IF (0 = bds_can_getDatabox(BDS_CAN_1_D, 1, DataboxData_au8[1], ADR(DataboxNumBytes_u8))) THEN
///  
///    (* Data in array DataboxData_au8 are valid and can be evaluated. *)
///	
///    (* The number of received bytes is stored in variable DataboxNumBytes_au8. *)
///  END_IF
///END
///
///============================================================================
{attribute 'external_name' := 'cmp_rts_bds_can_getDatabox'}
FUNCTION bds_can_getDatabox : UINT
VAR_INPUT
	///Indicates the CAN channel.Possible values are
	///    + BDS_CAN_1_D(0)
	///    + BDS_CAN_2_D(1)
	///    + BDS_CAN_3_D(2)
	///	+ BDS_CAN_4_D(3)
	chnl_e: bds_can_Chnl_te;
	///Receive databox number.
	///	
	///Each receive databox is numbered separately for each CAN channel.
	///
	///Value range: 1 .. n.
	///
	///n is the number of databoxes configured by easyConfig.
	databoxNum_u16: UINT;
	///Pointer to data array with at least 8 bytes.
	///	
	///The oldest data received by the configured databox is copied to this address. 
	data_pau8: POINTER TO USINT;
	///Number of bytes which are copied to data array data_pau8.
	numBytes_pu8: POINTER TO USINT;
END_VAR

END_FUNCTION

// Communication API/CAN/CAN legacy/API/bds_can_initRxDatabox
///This function initializes a CAN receive databox.
///
///=======
/// Remarks:
///=======
///    + The use of receive databoxes is optional!
///    + The number of required receive databoxes must be defined by easyConfig before using this function!
///    + Each receive databox has to be initialized before it can be used.
///    + The |GVL_can| is given for usage of defines.
///    + This API should be called once in Application
///
///----------
/// FFI:
///----------
///This API can be used in trusted partitions only. See Freedom from Interference (FFI) concept for more details.
///
///==================================================================		  			===================================================================================================
///Return value    								  									Description
///==================================================================		  			===================================================================================================
///0: BDS_CAN_ERR_NO_ERRORS_DU16														Function is called without errors. Receive databox was initialized successfully.
///9: BDS_CAN_ERR_DATABOXNUM_DU16														Invalid databox number.
///14: BDS_CAN_ERR_CHNL_DU16															Unknown CAN channel.
///15: BDS_CAN_ERR_ID_DU16																Invalid CAN identifier.
///16: BDS_CAN_ERR_FORMAT_DU16															Invalid message format.
///17: BDS_CAN_ERR_NUM_DATA_DU16														Invalid number of data bytes.
///55: BDS_CAN_ERR_OVERLAP_ADDR_DU16													Buffer overlaps with buffer registered already.
///60: BDS_CAN_ERR_INVALID_ADDR_DU16													NA.
///61: BDS_CAN_ERR_INVALID_ADDR_DU16													Invalid address (parameter buf_pas).Buffer length is zero.
///63: BDS_CAN_ERR_DATABOX_ID_EXIST_DU16												A databox with this identifier is initialised already.The new initialization will be not accepted.
///
///==================================================================		   			===================================================================================================
///=======
///Code Example:
///=======
///============================================================================
///PROGRAM PLC_PRG
///VAR
///	CAN_1_RX_DATABOX_1_BUF_LEN_DU8: UINT := 5;
///	can_1_RxDatabox_1_Buf_as: ARRAY[0..5] OF bds_can_DataboxData_ts;
///	flag: BOOL;
///	DataboxData_au8: ARRAY[0 .. 7] OF INT;
///	num_bytes:INT:=8;
///	count: UINT;
///	status_u16: UINT;
///END_VAR
///IF flag = FALSE THEN
///	status_u16 := bds_can_initRxDatabox(BDS_CAN_1_D, 1, 16#12, BDS_CAN_STD_DU8, 8, ADR(can_1_RxDatabox_1_Buf_as),CAN_1_RX_DATABOX_1_BUF_LEN_DU8,0);
///	bds_can_init(BDS_CAN_1_D, BDS_BAUD_500K_DU32);
///	flag:= TRUE;
///END_IF
///============================================================================
{attribute 'external_name' := 'cmp_rts_bds_can_initRxDatabox'}
FUNCTION bds_can_initRxDatabox : UINT
VAR_INPUT
	///Indicates the CAN channel.Possible values are
	///    + BDS_CAN_1_D(0)
	///    + BDS_CAN_2_D(1)
	///    + BDS_CAN_3_D(2)
	///	+ BDS_CAN_4_D(3)
	chnl_e: bds_can_Chnl_te;
	///Receive databox number.
	///	
	///Each receive databox is numbered separately for each CAN channel.
	///
	///Value range: 1 .. n.
	///
	///n is the number of databoxes configured by easyConfig. 
	databoxNum_u16: UINT;
	///Identifier of CAN message.
	///
	///Value range:
	///    - 16#000 .. 16#7FF (11-bit standard format)
	///    - 16#00000000 .. 16#1FFFFFFF (29-bit extented format)
	id_u32: UDINT;
	///Indicates the format of the CAN message.
	///
	///Value range:
	///
	///    - BDS_CAN_STD_DU8  (11-bit standard format)
	///    - BDS_CAN_EXD_DU8  (29-bit extented format)
	format_u8: USINT;
	///Number of bytes which can be received at maximum.
	///
	///Value range: 0 .. 8
	numBytes_u8: USINT;
	///Pointer to array of data type bds_can_DataboxData_ts.
	buf_pas: POINTER TO bds_can_DataboxData_ts;
	///Length of buffer array (that means number of CAN messages).
	///At least a buffer for 1 message is required.
	///
	///Value range: 1 .. n
	buf_len_u16: UINT;
	///
	///Pointer to a callback function of data type UINT which is called if a new message was received. If this callback function is used, then a receive buffer with a length of at least 1 message is mandatory.
	callback_pf: POINTER TO UINT;
END_VAR

END_FUNCTION

// Communication API/CAN/CAN legacy/API/bds_can_init
///The bds_can_init function does the following tasks:
///1. Re-initializes the baud rate of the CAN channel concerned.
///2. Starts the CAN channel. Re-initializes the CAN channel concerned following a bus off.
///
///=======
/// Remarks:
///=======
///    + The CAN channels are already initialized with the default baudrate by easyConfig.
///    + The current baudrate can be changed with this function.
///    + If an error occurs, channel is remaining in the default mode.
///    + Buffers and data boxes related to the CAN channel will not be cleared!
///    + This function also enables the CAN transceiver, if this feature is available for this CAN channel.
///    + If the CAN was initialized with this function then the sample point has the default value 80%. Other sample point values can be used with function bds_can_initxt .
///    + The |GVL_can| is given for usage of defines.
///    + This API should be called once in Application
///
///----------
/// FFI:
///----------
///This API can be used in trusted partitions only. See Freedom from Interference (FFI) concept for more details.
///
///==================================================================		  			===================================================================================================
///Return value    								  									Description
///==================================================================		  			===================================================================================================
///0: BDS_CAN_ERR_NO_ERRORS_DU16														Function is called without errors. Message data returned in msg_s are valid.
///1: BDS_CAN_ERR_UNKNOWN_BAUDRATE_DU16												Baud rate is not valid.
///14: BDS_CAN_ERR_CHNL_DU16															Unknown CAN channel.
///
///==================================================================		   			===================================================================================================
///
///=======
///Code Example:
///=======
///============================================================================
///
///PROGRAM PLC_PRG
///  VAR
///  
///  	flag: UINT;
///  END_VAR
///
///  (* re-initialize CAN channel 1 with 500KBaud *)
///  
///IF flag = FALSE THEN
///  bds_can_init(BDS_CAN_1_D, BDS_BAUD_500K_DU32);
///
///	flag:= TRUE;
///  
///END_IF
///
///============================================================================
{attribute 'external_name' := 'cmp_rts_bds_can_init'}
FUNCTION bds_can_init : UINT
VAR_INPUT
	///Indicates the CAN channel.Possible values are
	///    + BDS_CAN_1_D(0)
	///    + BDS_CAN_2_D(1)
	///    + BDS_CAN_3_D(2)
	///	+ BDS_CAN_4_D(3)
	chnl_e: bds_can_Chnl_te;
	///Indicates the baud rate.
	///	
	///Possible values:
	///    + BDS_BAUD_125K_DU32,
	///    + BDS_BAUD_250K_DU32,
	///    + BDS_BAUD_500K_DU32,
	///    + BDS_BAUD_1000K_DU32
	baudRate_u32: UDINT;
END_VAR

END_FUNCTION

// Communication API/CAN/CAN legacy/API/bds_can_initxt
///The bds_can_initxt function can be used optionally and alternatively to the function |bds_can_init|, if a specific sample point is required. It does the following tasks:
///
///1. Re-initializes the baud rate(s) of the CAN channel concerned.
///2. Starts the CAN channel. Re-initializes the CAN channel concerned following a bus off.
///
///=======
/// Remarks:
///=======
///	+ The CAN channels are already initialized with the default baud rate by easyConfig.
///	+ The current baud rate can be changed with this function.
///	+ If an error occurs, channel is remaining in the default mode.
///	+ Buffers and data boxes related to the CAN channel will not be cleared!
///	+ This function also enables the CAN transceiver, if this feature is available for this CAN channel.
///    + The |GVL_can| is given for usage of defines.
///    + This API should be called once in Application
///
///----------
/// FFI:
///----------
///This API can be used in trusted partitions only. See Freedom from Interference (FFI) concept for more details.
///
///==================================================================		  			===================================================================================================
///Return value    								  									Description
///==================================================================		  			===================================================================================================
///0: BDS_CAN_ERR_NO_ERRORS_DU16														Function is called without errors. Message data returned in msg_s are valid.
///1: BDS_CAN_ERR_UNKNOWN_BAUDRATE_DU16												Baud rate is not valid.
///2: BDS_CAN_ERR_SAMPLEPOINT_DU16														Sample point is not valid.
///3: BDS_CAN_ERR_FD_BAUDRATE_DU16														Data baud rate (in CAN FD mode) is not valid for this baud rate.
///14: BDS_CAN_ERR_CHNL_DU16															Unknown CAN channel.
///
///==================================================================		   			===================================================================================================
///
///=======
///Code Example:
///=======
///============================================================================
///
///PROGRAM PLC_PRG
///
///VAR
///
///	flag: UINT;
///
///END_VAR
///  
///IF flag = FALSE THEN
///
///  (* initialize CAN channel 1 in CAN standard mode with 250KBaud and a sample point with 85% *)
///  
///  bds_can_initxt(BDS_CAN_1_D, BDS_BAUD_250K_DU32, 85, 0);
///
///	flag:= TRUE;
///
///
///  (* ... *)
///  
///END
///
///============================================================================
{attribute 'external_name' := 'cmp_rts_bds_can_initxt'}
FUNCTION bds_can_initxt : UINT
VAR_INPUT
	///Indicates the CAN channel.Possible values are
	///    + BDS_CAN_1_D(0)
	///    + BDS_CAN_2_D(1)
	///    + BDS_CAN_3_D(2)
	///	+ BDS_CAN_4_D(3)
	chnl_e: bds_can_Chnl_te;
	///Indicates the (arbitration) baud rate.
	///
	///Possible values:
	///    + BDS_BAUD_125K_DU32
	///    + BDS_BAUD_250K_DU32
	///    + BDS_BAUD_500K_DU32
	///    + BDS_BAUD_1000K_DU32
	baudRate_u32: UDINT;
	///Indicates the sample point in %. The value = 0 sets the sample point on the same default value which is also used with the function bds_can_init.
	///
	///Possible values [in %]: 80, 85 or 0
	samplePoint_u8: USINT;
	///CAN FD mode is not yet supported.
	///
	///Possible values: 
	///Value = 0: CAN standard mode. 
	baudRateFd_u32: UDINT;
END_VAR

END_FUNCTION

// Communication API/CAN/CAN_FFI_API/bds_can_getDatabox_ffi
{attribute 'external_name' := 'cmp_rts_bds_can_getDatabox_ffi'}
FUNCTION bds_can_getDatabox_ffi : UINT
VAR_INPUT
	///Indicates the CAN channel.Possible values are
	///    + BDS_CAN_1_D(0)
	///    + BDS_CAN_2_D(1)
	///    + BDS_CAN_3_D(2)
	///	+ BDS_CAN_4_D(3)
	chnl_e: bds_can_Chnl_te;
	///Receive databox number.
	///	
	///Each receive databox is numbered separately for each CAN channel.
	///
	///Value range: 1 .. n.
	///
	///n is the number of databoxes configured by easyConfig.
	databoxNum_u16: UINT;
	///Pointer to data array with at least 8 bytes.
	///	
	///The oldest data received by the configured databox is copied to this address. 
	data_pau8: POINTER TO USINT;
	///Number of bytes which are copied to data array data_pau8.
	numBytes_pu8: POINTER TO USINT;
END_VAR

END_FUNCTION

// Communication API/CAN/CAN legacy/API/bds_can_getRxBufStatus
///This function returns the status of the Rx buffer of a CAN channel.
///
///=======
/// Remarks:
///=======
///    + The |GVL_can| is given for usage of defines.
///
///==================================================================		  			===================================================================================================
///Return value    								  									Description
///==================================================================		  			===================================================================================================
///>0																					Number of CAN messages in Rx buffer of the specified CAN channel which have been received.
///0																					Rx buffer is empty.
///-1																					Invalid CAN channel.
///5: BDS_CAN_FFI_ACCESS_ERROR_DU16														FFI API access error.
///==================================================================		   			===================================================================================================
///
///----------
/// FFI:
///----------
///This API can be used in trusted partitions. For untrusted partitions use |bds_can_getRxBufStatus_ffi|. See Freedom from Interference (FFI) concept for more details.
///
///=======
///Code Example:
///=======
///============================================================================
///
///PROGRAM appl_Task_1
///  VAR
///    numMsg_s32: DINT := 16#00;
///  END_VAR
/// 
///  numMsg_s32 := bds_can_getRxBufStatus(BDS_CAN_1_D);
///
///  IF (numMsg_s32 > 0) THEN
///  
///    (* RX buffer contains messages which can be read with bds_can_getData() *)
///	
///  END_IF
///END
///
///============================================================================
{attribute 'external_name' := 'cmp_rts_bds_can_getRxBufStatus'}
FUNCTION bds_can_getRxBufStatus : DINT
VAR_INPUT
	///Indicates the CAN channel.Possible values are
	///    + BDS_CAN_1_D(0)
	///    + BDS_CAN_2_D(1)
	///    + BDS_CAN_3_D(2)
	///	+ BDS_CAN_4_D(3)
	chnl_e: bds_can_Chnl_te;
END_VAR

END_FUNCTION

// Communication API/CAN/CAN_FFI_API/bds_can_getRxBufStatus_ffi
{attribute 'external_name' := 'cmp_rts_bds_can_getRxBufStatus_ffi'}
FUNCTION bds_can_getRxBufStatus_ffi : DINT
VAR_INPUT
	///Indicates the CAN channel.Possible values are
	///    + BDS_CAN_1_D(0)
	///    + BDS_CAN_2_D(1)
	///    + BDS_CAN_3_D(2)
	///	+ BDS_CAN_4_D(3)
	chnl_e: bds_can_Chnl_te;
END_VAR

END_FUNCTION

// Communication API/CAN/CAN legacy/API/bds_can_getStatus
///The status of a CAN interface can be read.
///
///=======
/// Remarks:
///=======
///    + This function mainly reads the status of the software CAN interface.
///    + CAN controller states like bus-off or error-passive can't be read with this function.
///    + If the CAN controller enters the bus-off state it will be restarted automatically by the BSW.
///    + Bus-off events can be detected by the application by means of a bus-off callback function.
///    + A bus-off callback function can be registered with function |bds_can_registerBusOffCallback|.
///    + The |GVL_can| is given for usage of defines.
///
///==================================================================		  			===================================================================================================
///Return value    								  									Description
///==================================================================		  			===================================================================================================
///0: BDS_CAN_STATE_UNINIT_DU16														UNINIT mode: CAN controller is not yet initialized after power on.
///1: BDS_CAN_STATE_STOPPED_DU16														STOPPED mode: CAN controller is halted and does not operate on the network. This state is reached e.g. due to function call |bds_can_stop|. The CAN controller can be activated again with |bds_can_start|.
///2: BDS_CAN_STATE_STARTED_DU16														STARTED mode: CAN controller is activated and in the full-operational mode.
///3: BDS_CAN_STATE_SLEEP_DU16															SLEEP mode: CAN controller is in sleep mode
///5: BDS_CAN_FFI_ACCESS_ERROR_DU16														FFI API access error.
///
///==================================================================		   			===================================================================================================
///
///----------
/// FFI:
///----------
///This API can be used in trusted partitions. For untrusted partitions use |bds_can_getStatus_ffi|. See Freedom from Interference (FFI) concept for more details.
///
///=======
///Code Example:
///=======
///============================================================================
///
///PROGRAM appl_Task_1
///  VAR
///    CAN_Status_u16: UINT := 16#00;
///  END_VAR
///
///   (* status of CAN channel BDS_CAN_1_D *)
///   CAN_Status_u16 := bds_can_getStatus(BDS_CAN_1_D);
///
///   IF (BDS_CAN_STATE_STARTED_DU16 <> CAN_Status_u16) THEN
///      (* e.g. restart CAN or error handling *)
///   END_IF
///END
///
///============================================================================
{attribute 'external_name' := 'cmp_rts_bds_can_getStatus'}
FUNCTION bds_can_getStatus : UINT
VAR_INPUT
	///Indicates the CAN channel.Possible values are
	///    + BDS_CAN_1_D(0)
	///    + BDS_CAN_2_D(1)
	///    + BDS_CAN_3_D(2)
	///	+ BDS_CAN_4_D(3)
	chnl_e: bds_can_Chnl_te;
END_VAR

END_FUNCTION

// Communication API/CAN/CAN legacy/API/bds_can_registerBusOffCallback
///With this function a callback function can be registered for each CAN channel, which is called if a can bus off occurred.
///
///=======
/// Remarks:
///=======
///    + Registering of this callback function is optional.
///    + Callback function must be defined within the application program.
///    + The |GVL_can| is given for usage of defines.
///
///----------
/// NOTICE:
///----------
///After a bus off event the CAN communication is recovered automatically by the BSW.
///
///----------
/// WARNING:
///----------
///
///This function should be called only once in the application.
///
///----------
/// FFI:
///----------
///This API can be used in trusted partitions only. See Freedom from Interference (FFI) concept for more details.
///
///==================================================================		  			===================================================================================================
///Return value    								  									Description
///==================================================================		  			===================================================================================================
///0: BDS_CAN_ERR_NO_ERRORS_DU16														Function is called without errors. Callback function was initialized successfully.
///14: BDS_CAN_ERR_CHNL_DU16															Unknown CAN channel.
///60: BDS_CAN_ERR_INVALID_ADDR_DU16													Invalid address (parameter func_pf).
///99: BDS_CAN_ERR_CFG_NOTALLOWED_DU16													Configuration is not allowed.
///
///==================================================================		   			===================================================================================================
///=======
///Code Example:
///=======
///============================================================================
///
///PROGRAM PLC_PRG
///
///  VAR
///	
///  END_VAR
///
///  
///IF flag = FALSE THEN
///
///	bds_can_registerBusOffCallback(BDS_CAN_1_D, can_1_BusOffCallback);
///
///	flag:= TRUE;
///
///END_IF
///
///FUNCTION can_1_BusOffCallback
///
///VAR
///
///	status_u16: UINT;
///	
///END_VAR
///
///============================================================================
///
{attribute 'external_name' := 'cmp_rts_bds_can_registerBusOffCallback'}
FUNCTION bds_can_registerBusOffCallback : UINT
VAR_INPUT
	///Indicates the CAN channel.Possible values are
	///    + BDS_CAN_1_D(0)
	///    + BDS_CAN_2_D(1)
	///    + BDS_CAN_3_D(2)
	///	+ BDS_CAN_4_D(3)
	chnl_e: bds_can_Chnl_te;
	///Pointer to a callback function of data type UINT which is called if a bus off occurs.
	func_pf: POINTER TO UINT;
END_VAR

END_FUNCTION

// Communication API/CAN/CAN legacy/API/bds_can_stop
///This function stops the specified CAN channel.
///
///=======
/// Remarks:
///=======
///    + The CAN channel is disabled and no transmit and receive operation are executed any more.
///    + The stopped CAN channel can be restarted by calling function |bds_can_start|.
///    + Data in CAN buffers (receive/send + databoxes) are not deleted! Transmit buffers can be reset with |bds_can_resetTxBuf|.
///    + This function also disables the CAN transceiver, if this feature is available for this CAN channel. 
///    + The |GVL_can| is given for usage of defines.
///
///----------
/// FFI:
///----------
///This API can be used in trusted partitions only. See Freedom from Interference (FFI) concept for more details.
///
///==================================================================		  			===================================================================================================
///Return value    								  									Description
///==================================================================		  			===================================================================================================
///0: BDS_CAN_ERR_NO_ERRORS_DU16														Function is called without errors. CAN channel was restarted successfully.
///14: BDS_CAN_ERR_CHNL_DU16															Unknown CAN channel.
///
///==================================================================		   			===================================================================================================
///
///=======
///Code Example:
///=======
///============================================================================
///
///PROGRAM appl_Task_1
///  VAR
///  
///  END_VAR
///
///  IF (<condition for CAN stop>) THEN
///    bds_can_stop(BDS_CAN_1_D);
///  END_IF
///END
///
///============================================================================
{attribute 'external_name' := 'cmp_rts_bds_can_stop'}
FUNCTION bds_can_stop : UINT
VAR_INPUT
	///Indicates the CAN channel.Possible values are
	///    + BDS_CAN_1_D(0)
	///    + BDS_CAN_2_D(1)
	///    + BDS_CAN_3_D(2)
	///	+ BDS_CAN_4_D(3)
	chnl_e: bds_can_Chnl_te;
END_VAR

END_FUNCTION

// Communication API/CAN/CAN legacy/API/bds_can_start
///This function restarts the specified CAN channel.
///
///=======
/// Remarks:
///=======
///    + This function can be used to restart the CAN channel after it had been stopped by calling |bds_can_stop|.
///    + Data in CAN buffers (receive/send + databoxes) are not deleted! Transmit buffers can be reset with |bds_can_resetTxBuf|.
///    + This function also enables the CAN transceiver, if this feature is available for this CAN channel. 
///    + The |GVL_can| is given for usage of defines.
///
///----------
/// FFI:
///----------
///This API can be used in trusted partitions only. See Freedom from Interference (FFI) concept for more details.
///
///==================================================================		  			===================================================================================================
///Return value    								  									Description
///==================================================================		  			===================================================================================================
///0: BDS_CAN_ERR_NO_ERRORS_DU16														Function is called without errors. CAN channel was restarted successfully.
///14: BDS_CAN_ERR_CHNL_DU16															Unknown CAN channel.
///
///==================================================================		   			===================================================================================================
///
///=======
///Code Example:
///=======
///============================================================================
///
///PROGRAM appl_Task_1
///  VAR
///  
///    CAN_Status_u16: UINT := 16#00;
///  END_VAR
///
///  (* check status of CAN channel 1 *)
///  
///  CAN_Status_u16 := bds_can_getStatus(BDS_CAN_1_D);
///
///  (* if CAN is not running then perform an automatic CAN restart *)
///  
///  IF (BDS_CAN_STATE_STARTED_DU16 <> CAN_Status_u16) THEN
///  
///    bds_can_start(BDS_CAN_1_D);
///	
///  END_IF
///END
///
///============================================================================
{attribute 'external_name' := 'cmp_rts_bds_can_start'}
FUNCTION bds_can_start : UINT
VAR_INPUT
	///Indicates the CAN channel.Possible values are
	///    + BDS_CAN_1_D(0)
	///    + BDS_CAN_2_D(1)
	///    + BDS_CAN_3_D(2)
	///	+ BDS_CAN_4_D(3)
	chnl_e: bds_can_Chnl_te;
END_VAR

END_FUNCTION

// Communication API/CAN/CAN legacy/API/bds_can_resetTxBuf
///This function resets the specified transmit buffer(s) for a CAN channel.
///
///=======
/// Remarks:
///=======
///    + The Tx buffer and/or the Tx databoxes can be reset.
///    + This function can be used after a |bds_can_stop| to delete all buffered messages before restarting the bus again with |bds_can_start|.
///    + The |GVL_can| is given for usage of defines.
///
///==================================================================		  			===================================================================================================
///Return value    								  									Description
///==================================================================		  			===================================================================================================
///0: BDS_CAN_ERR_NO_ERRORS_DU16														Function is called without errors. Message data returned in msg_s are valid.
///2: BDS_CAN_ERR_INV_BUF_TYPE_DU16													Invalid buffer type.
///1: BDS_CAN_ERR_CHNL_DU16															Unknown CAN channel.
///
///==================================================================		   			===================================================================================================
///
///----------
/// FFI:
///----------
///This API can be used in trusted partitions only. See Freedom from Interference (FFI) concept for more details.
///
///=======
///Code Example:
///=======
///============================================================================
///
///PROGRAM appl_Task_1
///  VAR
///  
///  END_VAR
///
///  (* Tx buffer and all Tx data boxes of CAN channel 1 will be reset *)
///  
///  bds_can_resetTxBuf(BDS_CAN_1_D, BDS_CAN_BUFTYPE_BUF_DU8 OR BDS_CAN_BUFTYPE_DATABOXES_DU8);
///
///  (* ... *)
///END
///
///============================================================================
{attribute 'external_name' := 'cmp_rts_bds_can_resetTxBuf'}
FUNCTION bds_can_resetTxBuf : UINT
VAR_INPUT
	///Indicates the CAN channel.Possible values are
	///    + BDS_CAN_1_D(0)
	///    + BDS_CAN_2_D(1)
	///    + BDS_CAN_3_D(2)
	///	+ BDS_CAN_4_D(3)
	chnl_e: bds_can_Chnl_te;
	///Indicates the buffer type:
	///
	///Bit coded value:
	///    + bit 0 = Tx buffer (BDS_CAN_BUFTYPE_BUF_DU8)
	///    + bit 1 = all Tx data boxes  (BDS_CAN_BUFTYPE_DATABOXES_DU8)
	///
	///Value range: 0 .. 3
	bufType_u8: USINT;
END_VAR

END_FUNCTION

// Communication API/CAN/CAN_FFI_API/bds_can_getStatus_ffi
{attribute 'external_name' := 'cmp_rts_bds_can_getStatus_ffi'}
FUNCTION bds_can_getStatus_ffi : UINT
VAR_INPUT
	///Indicates the CAN channel.Possible values are
	///    + BDS_CAN_1_D(0)
	///    + BDS_CAN_2_D(1)
	///    + BDS_CAN_3_D(2)
	///	+ BDS_CAN_4_D(3)
	chnl_e: bds_can_Chnl_te;
END_VAR

END_FUNCTION

